(* IEC 61131-3 sources: daoli-st-library/DL_Process (part 38) *)

(* ---- FB_DL_InlineCheckweighGauge.st ---- *)
(*==============================================================================
 * 组件名称 (Component)  : FB_DL_InlineCheckweighGauge
 * 所属子库 (Sublibrary) : DL_Process
 * 当前版本 (Version)    : 1.0.0
 * 兼容性 (Platform)     : CODESYS 3.5 / TwinCAT 3 / 汇川 InoProShop（纯标准元素，无方言）
 * 功能描述 (Function)   : 在线称重动态窗判据与 σ 控制图。逐件判欠重/超重（不平顺：平滑会
 *                         漏掉单件超重），滑动统计窗给均值与样本标准差（分母 n−1，n≥5 前置
 *                         保证防除零），满窗后才判 σ 越控制限；可选的 ±3σ 冲击剔除只影响
 *                         统计窗，不影响逐件判据。不做传感器标定、不做零点跟踪（另有专件）、
 *                         不做剔除机构驱动。
 * 溯源 (Origin)         : 道莅 clean-room 防御性实现
 * 本文件内含 (Contains) : TYPE E_DL_GaugeWin / FUNCTION_BLOCK FB_DL_InlineCheckweighGauge
 * 依赖 (Depends)        : 无（仅 Standard.library 的 SQRT / ABS / MIN）
 * 红线自检 (Redline)    : 无外部全局变量、无硬件地址直引 ｜ 全变量中英双语同行注释
 *                         公差与控制限判零防除零 ｜ 样本非有限即丢弃并计丢弃数 ｜ 标准差前置
 *                         n≥5 且分母 n−1 ｜ σ 仅满窗判 ｜ 枚举显式赋值 ｜ CASE 含 ELSE 兜底
 *                         ｜ 本件无定时器/沿实例，全部为周期算术，故无周期刷新项
 * 错误码表 (Codes)      : 16#0005_0444 就绪（窗口统计正常）
 *                         16#0005_0445 预留：本版不发码（下一轮区间起点，禁止回填）
 *                         16#0005_0446 故障级 组态非法（公差 ≤0、窗长 <5、σ 限 ≤0）
 *                         16#0005_0447 故障级 目标重量非有限（逐件判据停判，统计继续）
 *                         16#0005_0448 信息级 样本非有限已丢弃（计入丢弃数）
 * 修订历史 (Revision)   : 2026-11-17  v1.0.0  首版入库 · R28 · 阶段三批 4
 * 验收向量 (Acceptance) : 正向 目标 500 g、公差 ±5、10 件 500±1 → 均值 ≈500、σ ≈0.7、
 *                         无报警
 *                         反向 一件 508 g → bOver 单件置位、uRejectCnt 不增（非剔除开关）、
 *                         均值仍 ≈500；σ 升到 6 超控制限 2 → bSpcAlarm；样本给 NaN →
 *                         16#0005_0448 且丢弃数 +1；窗长给 3 → 16#0005_0446
 *============================================================================*)

(*-----------------------------------------------------------------------------
 * 枚举: E_DL_GaugeWin（归属本功能块，同文件发布，全库唯一定义）
 *----------------------------------------------------------------------------*)
TYPE E_DL_GaugeWin :
(
    eEmpty := 0,    // 空窗：尚无有效样本 / Empty window, no valid sample yet
    eFill  := 10,   // 填充中：样本数未满窗长 / Filling, the sample count is below the window length
    eFull  := 20,   // 满窗：均值与 σ 可信 / Full window, the mean and sigma are trustworthy
    eFault := 99    // 故障：组态非法 / Fault, the configuration is invalid
);
END_TYPE

FUNCTION_BLOCK FB_DL_InlineCheckweighGauge
VAR_INPUT
    bEnable        : BOOL := FALSE;       // 使能 / Enable
    bSampleValid   : BOOL := FALSE;       // 本拍有有效样本 / A valid sample is present in this scan
    fWeight_g      : REAL := 0.0;         // 件重 [g]，域 0~50000 / Piece weight in grammes, domain 0 to 50000
    fTarget_g      : REAL := 500.0;       // 目标重量 [g] / Target weight in grammes
    fTolUp_g       : REAL := 5.0;         // 上公差带 [g]，须 >0 / Upper tolerance in grammes, must be positive
    fTolLow_g      : REAL := 5.0;         // 下公差带 [g]，须 >0 / Lower tolerance in grammes, must be positive
    uWinSamples    : UINT := 10;          // 统计窗长 [个]，域 5~50 / Statistical window length, domain 5 to 50
    fSigmaLimit_g  : REAL := 2.0;         // σ 控制限 [g]，域 0.1~20 / Sigma control limit in grammes, domain 0.1 to 20
    bOutlierReject : BOOL := FALSE;       // ±3σ 冲击剔除开关 / Plus minus three sigma outlier rejection switch
END_VAR
VAR_OUTPUT
    fMeanOut_g     : REAL;                // 窗口均值 [g] / Window mean in grammes
    fSigmaOut_g    : REAL;                // 窗口标准差 [g] / Window standard deviation in grammes
    bUnder         : BOOL;                // 本件欠重（逐件判据） / This piece is underweight
    bOver          : BOOL;                // 本件超重（逐件判据） / This piece is overweight
    bSpcAlarm      : BOOL;                // σ 越控制限（满窗后才判） / Sigma above the control limit, judged on a full window only
    uRejectCnt     : UDINT;               // 剔除件数 [件]（±3σ 剔除） / Outlier rejection count
    uSpcCnt        : UDINT;               // SPC 越限次数 [次] / SPC limit violation count
    eErr           : UDINT;               // 错误码，段位 16#0005_xxxx / Error code in segment 16#0005_xxxx
END_VAR
VAR
    _eWin          : E_DL_GaugeWin := E_DL_GaugeWin.eEmpty; // 窗口相位 / Window phase
    _bInit         : BOOL := FALSE;       // 首扫标志，取非判定 / First-scan flag, tested negated
    _bCfgOk        : BOOL;                // 组态合法标志 / Configuration valid flag
    _bTgtOk        : BOOL;                // 目标有限标志 / Target finite flag
    _bSpcLatched   : BOOL := FALSE;       // SPC 报警锁存（单拍计数用） / SPC alarm latch for one-shot counting
    _uWinEff       : UINT := 10;          // 生效窗长（钳制后）[个] / Effective window length after clamping
    _uIdx          : UINT := 1;           // 环形写指针 / Circular write index
    _uFill         : UINT := 0;           // 已填样本数 [个] / Number of samples collected
    _fSum          : REAL := 0.0;         // 样本和 [g] / Sample sum
    _fMean         : REAL := 0.0;         // 窗口均值 [g] / Window mean
    _fMeanOut_g    : REAL := 0.0;         // 窗口均值中间量（出口映射源）[g] / Window mean intermediate, source of the outlet [g]
    _fVar          : REAL := 0.0;         // 样本方差 [g²] / Sample variance
    _afWin         : ARRAY[1..50] OF REAL; // 样本环形窗 [g] / Sample ring buffer
    _iLoop         : INT;                 // 统计循环索引 / Statistical loop index
    _iGuard        : INT;                 // 防死循环计数器 / Loop guard counter
END_VAR
VAR CONSTANT
    DL_CW_READY    : UDINT := 16#0005_0444;  // 就绪码 / Ready code
    DL_CW_CFG_BAD  : UDINT := 16#0005_0446;  // 故障级组态非法码 / Fault code for bad configuration
    DL_CW_TGT_BAD  : UDINT := 16#0005_0447;  // 故障级目标非有限码 / Fault code for a non-finite target
    DL_CW_SKIP     : UDINT := 16#0005_0448;  // 信息级样本丢弃码 / Info code for a discarded sample
    DL_CW_WIN_LO   : UINT := 5;              // 窗长下限 [个] / Window length lower bound
    DL_CW_WIN_HI   : UINT := 50;             // 窗长上限 [个] / Window length upper bound
    DL_CW_SIG_LO   : REAL := 0.1;            // σ 控制限下限 [g] / Sigma limit lower bound
    DL_CW_SIG_HI   : REAL := 20.0;           // σ 控制限上限 [g] / Sigma limit upper bound
    DL_CW_LOOP_MAX : INT := 60;              // 循环保护上限 / Loop guard bound
    DL_CW_EPS      : REAL := 1.0E-6;         // 浮点判零容差 / Float zero tolerance
END_VAR

// 段 1｜输出与单拍标志预置
bUnder := FALSE;                                    // 欠重预清 / Underweight pre-cleared
bOver := FALSE;                                     // 超重预清 / Overweight pre-cleared
bSpcAlarm := FALSE;                                 // SPC 报警预清 / SPC alarm pre-cleared
eErr := 0;                                          // 错误码预清 / Error code pre-cleared

// 段 2｜首扫初始化（判据取非，R19）
IF NOT _bInit THEN
    _afWin[1] := 0.0;                               // 环形窗首元素预置 [g] / Ring buffer first element pre-set
    _eWin := E_DL_GaugeWin.eEmpty;                  // 窗口相位起点 / Window phase starts empty
    _bInit := TRUE;                                 // 首扫只做一次 / The first scan runs once
END_IF

// 段 3｜组态闸（公差与控制限判零防除零；窗长 <5 使 σ 不可信）
_bCfgOk := (fTolUp_g > 0.0) AND (fTolLow_g > 0.0)
        AND NOT ((fSigmaLimit_g <> fSigmaLimit_g) OR ((fSigmaLimit_g - fSigmaLimit_g) <> (fSigmaLimit_g - fSigmaLimit_g)))
        AND (fSigmaLimit_g >= DL_CW_SIG_LO) AND (fSigmaLimit_g <= DL_CW_SIG_HI)
        AND (uWinSamples >= DL_CW_WIN_LO) AND (uWinSamples <= DL_CW_WIN_HI);
_bTgtOk := NOT ((fTarget_g <> fTarget_g) OR ((fTarget_g - fTarget_g) <> (fTarget_g - fTarget_g)));
IF NOT _bCfgOk THEN
    eErr := DL_CW_CFG_BAD;                          // 故障级：组态非法 / Fault, bad configuration
    _eWin := E_DL_GaugeWin.eFault;
ELSE
    _uWinEff := uWinSamples;                        // 采用组态窗长 [个] / Use the configured window length
END_IF
IF NOT _bTgtOk THEN
    eErr := DL_CW_TGT_BAD;                          // 故障级：目标非有限（逐件判据停判） / Fault, the target is not finite
END_IF

// 段 4｜逐件判据（不平顺，单件即判；目标不可读时停判）
IF bEnable AND bSampleValid AND _bTgtOk THEN
    IF (fWeight_g <> fWeight_g) OR ((fWeight_g - fWeight_g) <> (fWeight_g - fWeight_g)) THEN
        eErr := DL_CW_SKIP;                         // 信息级：样本非有限，丢弃 / Info, the sample is not finite and is discarded
        uRejectCnt := uRejectCnt + 1;               // 丢弃计数 +1 [件] / Discard count incremented
    ELSE
        IF fWeight_g < (fTarget_g - fTolLow_g) THEN
            bUnder := TRUE;                         // 本件欠重 / This piece is underweight
        END_IF
        IF fWeight_g > (fTarget_g + fTolUp_g) THEN
            bOver := TRUE;                          // 本件超重 / This piece is overweight
        END_IF
        // 冲击剔除（±3σ，仅满窗且开关有效时；剔除只影响统计窗）
        IF bOutlierReject AND (_uFill >= DL_CW_WIN_LO) AND (fSigmaOut_g > DL_CW_EPS) THEN
            IF ABS(fWeight_g - _fMean) > (3.0 * fSigmaOut_g) THEN
                uRejectCnt := uRejectCnt + 1;       // ±3σ 剔除 +1 [件] / Outlier rejected
            ELSE
                _fSum := _fSum - _afWin[_uIdx];                 // 换出最旧样本 [g] / Remove the oldest sample
                _afWin[_uIdx] := fWeight_g;                     // 写入新样本 [g] / Insert the new sample
                _fSum := _fSum + fWeight_g;                     // 样本和更新 [g] / Update the sum
                _uIdx := _uIdx + 1;
                IF _uIdx > _uWinEff THEN
                    _uIdx := 1;                                 // 环形回卷 / Ring wrap
                END_IF
                IF _uFill < _uWinEff THEN
                    _uFill := _uFill + 1;                       // 已填样本数 +1 [个] / Sample count incremented
                END_IF
            END_IF
        ELSE
            _fSum := _fSum - _afWin[_uIdx];                     // 换出最旧样本 [g] / Remove the oldest sample
            _afWin[_uIdx] := fWeight_g;                         // 写入新样本 [g] / Insert the new sample
            _fSum := _fSum + fWeight_g;                         // 样本和更新 [g] / Update the sum
            _uIdx := _uIdx + 1;
            IF _uIdx > _uWinEff THEN
                _uIdx := 1;                                     // 环形回卷 / Ring wrap
            END_IF
            IF _uFill < _uWinEff THEN
                _uFill := _uFill + 1;                           // 已填样本数 +1 [个] / Sample count incremented
            END_IF
        END_IF
    END_IF
END_IF

// 段 5｜均值与样本标准差（分母 n−1，n≥5 前置保证防除零）
IF _uFill > 0 THEN
    _fMean := _fSum / UINT_TO_REAL(_uFill);         // 窗口均值 [g] / Window mean
END_IF
_fMeanOut_g := _fMean;                              // 均值出口 [g] / Mean output
_fVar := 0.0;                                       // 方差清零 [g²] / Variance reset
IF _uFill >= DL_CW_WIN_LO THEN
    _iLoop := 1;
    _iGuard := 0;
    WHILE (_iLoop <= UINT_TO_INT(_uWinEff)) AND (_iGuard < DL_CW_LOOP_MAX) DO
        _fVar := _fVar + ((_afWin[_iLoop] - _fMean) * (_afWin[_iLoop] - _fMean));   // 偏差平方累加 [g²] / Squared deviation accumulated
        _iLoop := _iLoop + 1;
        _iGuard := _iGuard + 1;                     // 防死循环计数 / Loop guard incremented
    END_WHILE
    _fVar := _fVar / UINT_TO_REAL(_uWinEff - 1);    // 样本方差（分母 n−1）[g²] / Sample variance with n minus one
    fSigmaOut_g := SQRT(_fVar);                     // 样本标准差 [g] / Sample standard deviation
ELSE
    fSigmaOut_g := 0.0;                             // 样本不足：σ 记 0（不参与判据） / Not enough samples, sigma reported as zero
END_IF

// 段 6｜σ 控制图（仅满窗判；越限只在锁存沿计数一次）
IF (_uFill >= _uWinEff) AND (_uWinEff >= DL_CW_WIN_LO) THEN
    IF fSigmaOut_g > fSigmaLimit_g THEN
        bSpcAlarm := TRUE;                          // σ 越控制限 / Sigma above the control limit
        IF NOT _bSpcLatched THEN
            uSpcCnt := uSpcCnt + 1;                 // 越限次数 +1（沿计数）[次] / Violation count incremented on the edge
            _bSpcLatched := TRUE;
        END_IF
    ELSE
        _bSpcLatched := FALSE;                      // 回限内：锁存解除 / Back inside the limit, the latch is released
    END_IF
END_IF

// 段 7｜窗口相位映射（ENUM + CASE + ELSE 兜底）
CASE _eWin OF
    E_DL_GaugeWin.eEmpty:
        IF _uFill > 0 THEN
            _eWin := E_DL_GaugeWin.eFill;           // 有样本：进入填充 / Samples exist, go filling
        END_IF
    E_DL_GaugeWin.eFill:
        IF _uFill >= _uWinEff THEN
            _eWin := E_DL_GaugeWin.eFull;           // 满窗 / Window full
        END_IF
    E_DL_GaugeWin.eFull:
        IF _uFill < _uWinEff THEN
            _eWin := E_DL_GaugeWin.eFill;           // 窗被重置 / The window was reset
        END_IF
    E_DL_GaugeWin.eFault:
        IF _bCfgOk THEN
            _eWin := E_DL_GaugeWin.eEmpty;          // 组态修正：回空窗 / Configuration fixed, back to empty
        END_IF
        eErr := DL_CW_CFG_BAD;                      // 故障级：组态非法保持 / Fault, the configuration error is held
    ELSE
        // 非法相位兜底（故障级）
        eErr := DL_CW_CFG_BAD;
        _eWin := E_DL_GaugeWin.eFault;
END_CASE
IF eErr = 0 THEN
    eErr := DL_CW_READY;                            // 无事件回就绪码 / Ready code when nothing else applies
END_IF
END_FUNCTION_BLOCK

(* ---- FB_DL_InvInsulTestSeq.st ---- *)
(*
  FB_DL_InvInsulTestSeq  —  逆变器绝缘测试加压-保持-泄放联锁顺控 / Inverter insulation test sequence with discharge interlock
  分类 Category : DL_Process
  码位 Code     : 16#06_0_98
  版本 Version  : 1.0.0
  溯源 Source   : ISA-88 相模型语义借鉴 · clean-room 实现，仅借分类/参数域/命名，未复制源码
  功能 Function : 1) 加压-保持-泄放三态顺控（复用 FB_DL_InterlockMatrix 联锁前置）；
                  2) 加压中急停立即转泄放相（安全侧打断）；
                  3) 泄放未确认前禁放行下工序；相完成仅在泄放反馈确认后置位。
  边界 Boundary : ① 泄放未确认前禁放行下工序（安全侧默认，bTestOk 不置位）；
                  ② 加压中急停立即转泄放相（打断优先级最高）；
                  ③ 各相超时独立 TON 升级；
                  ④ 测试电压反馈无效判「不可判」而非 OK；
                  ⑤ 输出三行同向：相状态 → 测试结论 → 联锁出口。
  依赖 Depends  : FB_DL_InterlockMatrix × 1（联锁前置，每拍无条件调用）

  码表 Error codes（本件子码步进 16#30 · 本格 98 与既有 9X 子码段冲突，错位至 C8/D8 避让）:
    16#0002_06C8 故障级：组态非法（任一相时长 <= 0 / 电压门限 <= 0）
    16#0002_06D8 故障级：相超时（加压/保持/泄放任一相在限时内未完成，锁存需复位）
    16#0002_06B8 信息级：电压反馈无效判不可判 / 泄放未确认不放行（不置 bError）
*)

TYPE E_DL_IitPhase :
(
    eIdle       := 0,  // 空闲 / Idle
    ePressurize := 10, // 加压相 / HV apply phase
    eHold       := 20, // 保持相 / Hold phase
    eDischarge  := 30, // 泄放相 / Discharge phase
    eDone       := 40, // 测试完成（泄放已确认）/ Test done, discharge confirmed
    eFault      := 90  // 超时/联锁故障锁定 / Timeout or interlock fault locked
);
END_TYPE

FUNCTION_BLOCK FB_DL_InvInsulTestSeq
VAR_INPUT
    bTestCmd      : BOOL;                           // 测试启动命令 / Test start command
    bEStop        : BOOL;                           // 急停（加压/保持相打断转泄放）/ Emergency stop
    bVoltFbOk     : BOOL;                           // 电压反馈有效前置 / Voltage feedback valid flag
    fVoltFb       : REAL;                           // 测试电压反馈 [V] / Test voltage feedback [V]
    fVoltSp       : REAL := 1000.0;                 // 测试电压设定 [V]，域 > 0 / Test voltage setpoint [V]
    fVoltWinV     : REAL := 50.0;                   // 保持相电压窗半宽 [V]，域 > 0 / Hold voltage window [V]
    bDischargeFb  : BOOL;                           // 泄放反馈（残压低于安全值）/ Discharge feedback, residual below safe
    bReset        : BOOL;                           // 复位，上升沿清故障 / Reset, clears fault
    tApplyMax     : TIME := T#10S;                  // 加压相限时 [s]，域 > 0 / Apply phase timeout
    tHoldMax      : TIME := T#5S;                   // 保持相限时 [s]，域 > 0 / Hold phase timeout
    tDischMax     : TIME := T#30S;                  // 泄放相限时 [s]，域 > 0 / Discharge phase timeout
    fEps          : REAL := 1.0E-6;                 // 浮点判零容差 [1] / Floating zero tolerance
END_VAR
VAR_OUTPUT
    bApplyHv      : BOOL;                           // 加压出口 / HV apply output
    bDischargeCmd : BOOL;                           // 泄放命令出口 / Discharge command output
    bTestOk       : BOOL;                           // 测试结论（仅在泄放确认后置位）/ Test verdict, only after discharge confirmed
    bInterlock    : BOOL;                           // 联锁出口（TRUE = 允许加压）/ Interlock output
    bIndeterminate: BOOL;                           // 不可判标志（反馈无效）/ Indeterminate flag
    bError        : BOOL;                           // 故障标志，与故障级码配对 / Fault flag
    uErrorId      : UDINT;                          // 事件码，0 = 无事件 / Event code
    eStateOut     : E_DL_IitPhase;                  // 状态机当前态，段尾单点映射 / Phase mapped at tail
END_VAR
VAR
    _eState       : E_DL_IitPhase := E_DL_IitPhase.eIdle;  // 内部状态 / Internal state
    fbIlk         : FB_DL_InterlockMatrix;          // 联锁矩阵实例（无条件调用）/ Interlock matrix instance
    rtrStart      : R_TRIG;                         // 启动沿 / Start edge
    rtrReset      : R_TRIG;                         // 复位沿 / Reset edge
    tonApply      : TON;                            // 加压相超时（独立 TON）/ Apply timeout
    tonHold       : TON;                            // 保持相超时 / Hold timeout
    tonDisch      : TON;                            // 泄放相超时 / Discharge timeout
    abCondOk      : ARRAY[0..15] OF BOOL;           // 联锁条件表 / Interlock condition table
    auInvertMask  : WORD;                           // 取反掩码 / Invert mask
    auTripMask    : WORD;                           // 停机级掩码 / Trip-class mask
    bCfgOk        : BOOL;                           // 组态合法标志 / Configuration valid
    bVoltOk       : BOOL;                           // 电压反馈本拍有效 / Voltage feedback valid
    bVoltInWin    : BOOL;                           // 保持相电压在窗 / Hold voltage in window
    bIlkPermit    : BOOL;                           // 联锁放行 / Interlock permit
    uFault        : UDINT;                          // 锁存故障码 / Latched fault code
    uInfo         : UDINT;                          // 信息级码 / Information code
END_VAR

(* === 段 0 · 实例刷新 === *)
rtrStart(CLK := bTestCmd);                        // 每拍刷新启动沿
rtrReset(CLK := bReset);                          // 每拍刷新复位沿

(* === 段 1 · 组态闸 === *)
bCfgOk := (TIME_TO_REAL(tApplyMax) > fEps) AND (TIME_TO_REAL(tHoldMax) > fEps)
          AND (TIME_TO_REAL(tDischMax) > fEps)    // 三相时长正域
          AND (fVoltSp > fEps) AND (fVoltWinV > fEps)   // 电压设定与窗正域
          AND (fVoltSp = fVoltSp) AND (fVoltWinV = fVoltWinV);  // NaN 自反
IF NOT bCfgOk THEN
    uFault := 16#0002_06C8;                       // 故障级：组态非法
END_IF
IF rtrReset.Q AND bCfgOk THEN
    uFault := 16#0000;                            // 复位沿清锁存（解除路径可达）
END_IF
uInfo := 16#0000;                                 // 信息码每拍清零

(* === 段 2 · 相超时定时器（独立 TON，相离开即断输入，R40）=== *)
tonApply(IN := (_eState = E_DL_IitPhase.ePressurize), PT := tApplyMax);   // 加压相超时
tonHold(IN := (_eState = E_DL_IitPhase.eHold), PT := tHoldMax);           // 保持相超时
tonDisch(IN := (_eState = E_DL_IitPhase.eDischarge), PT := tDischMax);    // 泄放相超时
IF tonApply.Q OR tonHold.Q OR tonDisch.Q THEN
    uFault := 16#0002_06D8;                       // 故障级：任一相超时（锁存，非死等）
END_IF

(* === 段 3 · 联锁矩阵（无条件调用：急停未触发 + 电压反馈有效 + 复位态）=== *)
abCondOk[0] := NOT bEStop;                        // 条件 0 = 急停未触发
abCondOk[1] := bVoltFbOk;                         // 条件 1 = 电压反馈有效
abCondOk[2] := bDischargeFb OR (_eState = E_DL_IitPhase.eIdle);   // 条件 2 = 初始无残压或空闲态
auInvertMask := 16#0000;                          // 不取反
auTripMask := 16#0007;                            // 三条件均停机级
fbIlk(abConditionOk := abCondOk,                  // 条件表
      auInvertMask := auInvertMask,               // 取反掩码
      auTripMask := auTripMask,                   // 停机级掩码
      bEnable := TRUE,                            // 矩阵恒使能（安全联锁语义由条件表与停机级掩码承载）
      bReset := rtrReset.Q);                      // 复位沿透传
bIlkPermit := fbIlk.bPermitToRun;                 // 联锁放行
bInterlock := bIlkPermit;                         // 联锁出口

(* === 段 4 · 电压反馈域闸与保持窗判定 === *)
bVoltOk := bVoltFbOk AND (fVoltFb = fVoltFb) AND (fVoltFb >= 0.0) AND (fVoltFb < 1.0E30);  // NaN 自反 + 非负域
bVoltInWin := bVoltOk AND (ABS(fVoltFb - fVoltSp) <= fVoltWinV + fEps);   // 保持相电压在窗
IF (_eState = E_DL_IitPhase.eHold) AND (NOT bVoltOk) THEN
    uInfo := 16#0002_06B8;                        // 信息级：电压反馈无效判不可判
END_IF
bIndeterminate := (NOT bVoltOk) AND ((_eState = E_DL_IitPhase.eHold)
                    OR (_eState = E_DL_IitPhase.ePressurize));   // 不可判标志（非 OK）

(* === 段 5 · 主状态机（ENUM + CASE，含 ELSE 兜底）=== *)
CASE _eState OF
E_DL_IitPhase.eIdle :
    bTestOk := FALSE;                             // 空闲未完成
    IF uFault <> 16#0000 THEN
        _eState := E_DL_IitPhase.eFault;          // 故障优先
    ELSIF rtrStart.Q AND bIlkPermit AND bCfgOk THEN
        _eState := E_DL_IitPhase.ePressurize;     // 联锁放行才进加压相
    END_IF

E_DL_IitPhase.ePressurize :
    bApplyHv := bIlkPermit AND (uFault = 16#0000);   // 加压出口（联锁+无故障门控）
    bDischargeCmd := FALSE;                       // 加压相不出泄放命令
    IF bEStop THEN
        _eState := E_DL_IitPhase.eDischarge;      // 急停立即转泄放相（打断优先级最高）
    ELSIF uFault <> 16#0000 THEN
        _eState := E_DL_IitPhase.eFault;          // 超时转故障
    ELSIF bVoltInWin THEN
        _eState := E_DL_IitPhase.eHold;           // 电压进窗转保持相
    END_IF

E_DL_IitPhase.eHold :
    bApplyHv := TRUE;                             // 保持相维持加压
    bDischargeCmd := FALSE;                       // 保持相不出泄放命令
    IF bEStop THEN
        _eState := E_DL_IitPhase.eDischarge;      // 急停立即转泄放相
    ELSIF uFault <> 16#0000 THEN
        _eState := E_DL_IitPhase.eFault;          // 超时转故障
    ELSIF tonHold.Q THEN
        _eState := E_DL_IitPhase.eDischarge;      // 保持时限到转泄放相（正常流程）
    END_IF

E_DL_IitPhase.eDischarge :
    bApplyHv := FALSE;                            // 泄放相撤加压
    bDischargeCmd := TRUE;                        // 泄放命令保持
    IF uFault <> 16#0000 THEN
        _eState := E_DL_IitPhase.eFault;          // 泄放超时转故障
    ELSIF bDischargeFb AND (NOT bEStop) THEN
        bTestOk := TRUE;                          // 泄放反馈确认：相完成仅此时置位
        _eState := E_DL_IitPhase.eDone;           // 转完成相
    ELSE
        uInfo := 16#0002_06B8;                    // 信息级：泄放未确认不放行
    END_IF

E_DL_IitPhase.eDone :
    bApplyHv := FALSE;                            // 完成相撤加压
    bDischargeCmd := FALSE;                       // 完成相撤泄放命令
    bTestOk := TRUE;                              // 结论保持（防同拍抹除）
    IF rtrStart.Q THEN
        bTestOk := FALSE;                         // 新启动沿重开
        _eState := E_DL_IitPhase.ePressurize;     // 回加压相
    END_IF

E_DL_IitPhase.eFault :
    bApplyHv := FALSE;                            // 故障相撤加压
    bDischargeCmd := TRUE;                        // 故障安全侧：泄放命令保持
    bTestOk := FALSE;                             // 故障不出结论
    IF uFault = 16#0000 THEN
        _eState := E_DL_IitPhase.eIdle;           // 解锁回空闲
    END_IF

ELSE
    _eState := E_DL_IitPhase.eFault;              // 非法状态拦截
    uFault := 16#0002_06C8;                       // 故障级：相 ID 越界复用组态码段
END_CASE

(* === 段 6 · 输出映射 === *)
bError := (uFault <> 16#0000);                    // 故障标志仅由故障级码置位（R45 配对）
IF bError THEN
    uErrorId := uFault;                           // 故障级优先上报
ELSE
    uErrorId := uInfo;                            // 否则上报信息级码
END_IF
eStateOut := _eState;                             // 输出枚举段尾单点映射（N2 规则）
END_FUNCTION_BLOCK

(* ---- FB_DL_IvCurveScan.st ---- *)
(*
  FB_DL_IvCurveScan  —  IV 曲线扫描与特征点提取（Voc / Isc / FF + 扫描窗） / IV curve scan with Voc, Isc and fill-factor extraction inside a scan window
  分类 Category : DL_Process
  版本 Version  : 1.0.1
  来源 Source   : roadmap-pv-p1 — 光伏组件 IV 扫描测试工站真缺口
  溯源 Origin   : 道莅 clean-room 实现；Voc/Isc/Pmax/FF 为公开光伏特性参数定义式，未复制任何源码行
  功能 Function : 1) 扫描窗 eScan 内逐周期摄取 (fVmeasV, fImeasA) 采样：Voc = 电压最大值、
                  Isc = 电流最大值、Pmax = max(V×I) 功率最大值、nSample 采样计数；
                  2) 段 0 每拍单次求解 FF = Pmax/(Voc×Isc)，内核为纯计算子函数
                  FC_DL_IvFillFactorCalc（分母 <= 1.0E-9 返回 -1.0 哨兵，不饱和、不置 0），
                  判据与出口共用同一当拍量 _fFfPu，全件不存在同一子函数同参二次调用；
                  3) FF 低于 fFfMinPu 判组件异常（归因 eFfLow）；
                  4) 故障级单码 03A2，归因由 eCause 独立成员承载（R190）；
                  5) 信息级 04CA = 扫描完成沿；6) 解除式全当拍量（R240）。
  接口 Interface: 输入逐样电压/电流/扫描窗/最小采样数/FF 下限/电压量程；输出 Voc/Isc/Pmax/FF/采样数/码
  边界 Boundary : ① 组态闸：tScan <= T#0S、nSampleMin = 0、fFfMinPu <= 0.0、fVmaxV <= 0.0
                  任一成立 → 03A2 锁存；fFfMinPu / fVmaxV 同时做 NaN 自反判，否则 NaN 参与
                  `<= 0.0` 判据恒假 → 组态闸与「FF 越下限」判据双双静默失效；
                  ② 非有限输入（NaN 自反 + Inf 差值自减双判）→ 03A2 锁存且该样点不参与极值更新；
                  ③ 除零防护在子函数内前置判（分母非法返回 -1.0 哨兵，不饱和、不置 0）；
                  ④ 采样极值仅扫峰不回落（扫描窗内单调保持），窗口结束由 TON 单点置位；
                  ⑤ 扫描 TON / R_TRIG 段 0 无条件周期调用，IN 由相位派生；
                  ⑥ 零全局耦合（无 GVL / 无 VAR_EXTERNAL / 无直接物理地址访问）；
                  ⑦ 复位沿作用域（R283 返修）：eFault 相内 = 清故障三件 + 净重装窗内量并回 eIdle；
                  非故障相 = 仅清故障锁存三件，窗内量与相位一律不动；窗内量唯一重置点 =
                  eIdle→eScan 迁移（段 5），保证「复位不清窗」与「tonScan 不重装」自洽；
                  ⑧ 〔例外〕NaN 自反判 [x <> x] 与 Inf 差值自减判 [(x-x) <> (x-x)] 是浮点判等
                  禁令的唯一合法例外（R79），只许用于「非有限检测」；机检 G6 已对自反式加白名单。
  依赖 Depends  : Standard.library（TON / R_TRIG）
  码表 Error codes（Process 段 0005，故障窗口 03A2 / 信息窗口 04CA）:
    16#0005_03A2 故障级：IV 扫描故障总码（组态非法 / 输入非有限 / 采样数不足 / FF 越下限），
                 锁存至 bReset 上升沿；归因见 eCause，不新增码位（派单硬约束单码）
    16#0005_04CA 信息级：扫描完成沿（进入 eDone 单拍）
  修订历史 Revision :
    2026-11-19  v1.0.0  R43 首版（批次 2 · 序号 6）
    2026-11-19  v1.0.1  R45 返修（R283）：复位沿按相分域，非故障相不再清窗内极值与采样计数
                        （曾致 eScan 中复位后半窗从零累积、与 tonScan 不重装自相矛盾）；
                        FF 计算上移段 0 单次求解 _fFfPu，段 3 判据与 eEval 相改读当拍量，
                        删除同一 FC 同参双调用；出口 fFfPu 恒等 _fFfPu，消除 eDone 相 FF 恒 0；
                        组态闸补 NaN 自反判；边界新增⑦⑧；引脚契约零变更（PATCH）
*)

TYPE E_DL_IvsState :
(
    eIdle  := 0,      // 未使能待启动 / Idle, waiting start
    eScan  := 10,     // 扫描窗内逐样摄取 / Sampling inside scan window
    eEval  := 20,     // 特征点求解与判据 / Feature evaluation
    eDone  := 50,     // 扫描完成 / Done
    eFault := 90      // 故障锁存相 / Fault latched phase
);
END_TYPE

TYPE E_DL_IvsCause :
(
    eNone       := 0, // 无故障成因 / No cause
    eCfgIllegal := 1, // 组态非法 / Illegal configuration
    eNonFinite  := 2, // 输入非有限 / Non-finite input
    eSampleFew  := 3, // 采样数不足 / Too few samples
    eFfLow      := 4  // FF 越下限（含分母不可计算时 FF 不可达下限） / Fill factor below limit
);
END_TYPE

FUNCTION FC_DL_IvFillFactorCalc : REAL
VAR_INPUT
    fPmaxW : REAL;    // 最大功率 [W] / Maximum power
    fVocV  : REAL;    // 开路电压 [V] / Open-circuit voltage
    fIscA  : REAL;    // 短路电流 [A] / Short-circuit current
END_VAR
(* 纯计算子函数：FF = Pmax / (Voc × Isc)；分母 <= 1.0E-9 返回 -1.0 哨兵（不饱和、不置 0） *)
IF (fVocV <= 1.0E-9) OR (fIscA <= 1.0E-9) THEN      // 除零前置判（分母正域检查） / Divide-by-zero guard
    FC_DL_IvFillFactorCalc := -1.0;                 // 哨兵：分母非法 / Sentinel for invalid denominator
ELSE
    FC_DL_IvFillFactorCalc := fPmaxW / (fVocV * fIscA);   // 填充因子（无量纲） / Fill factor
END_IF
END_FUNCTION

FUNCTION_BLOCK FB_DL_IvCurveScan
VAR_INPUT
    fVmeasV      : REAL := 0.0;       // 逐样电压 [V] / Per-sample voltage
    fImeasA      : REAL := 0.0;       // 逐样电流 [A] / Per-sample current
    tScan        : TIME := T#2S;      // 扫描窗时长 [ms]，域 > 0 / Scan window duration
    nSampleMin   : UDINT := 20;       // 最小采样点数 [点]，域 > 0 / Minimum sample count
    fFfMinPu     : REAL := 0.60;      // FF 下限 [p.u.]，域 > 0 / Fill factor lower limit
    fVmaxV       : REAL := 60.0;      // 电压量程上限 [V]，域 > 0 / Voltage range limit
    bStart       : BOOL := FALSE;     // 启动命令（电平）[-] / Start command
    bReset       : BOOL := FALSE;     // 复位命令，上升沿清故障 [-] / Reset edge
END_VAR
VAR_OUTPUT
    eState       : E_DL_IvsState;     // 状态出口，段 6 单点映射 / State outlet
    eCause       : E_DL_IvsCause;     // 故障成因出口（R190） / Fault cause outlet
    fVocV        : REAL;              // 开路电压 [V] / Open-circuit voltage
    fIscA        : REAL;              // 短路电流 [A] / Short-circuit current
    fPmaxW       : REAL;              // 最大功率 [W] / Maximum power
    fFfPu        : REAL;              // 填充因子 [p.u.] / Fill factor
    nSampleCount : UDINT;             // 本次扫描采样点数 [点] / Sample count
    bCycleDone   : BOOL;              // 扫描完成标志 [-] / Scan done flag
    bError       : BOOL;              // 故障锁存标志 [-] / Fault latch flag
    nErrId       : UDINT;             // 事件码，0 = 无事件 / Event code
END_VAR
VAR
    _eState      : E_DL_IvsState := E_DL_IvsState.eIdle;   // 内部相位（CASE 唯一写入目标） / Internal phase
    _eCause      : E_DL_IvsCause := E_DL_IvsCause.eNone;   // 故障成因锁存（锁存量） / Latched cause
    tonScan      : TON;               // 扫描窗计时，每周期无条件调用 / Scan window timer
    rtReset      : R_TRIG;            // 复位沿实例，每周期无条件调用 / Reset edge
    _fVocV       : REAL;              // 扫描期电压极值（窗内保持） / Voltage peak held in window
    _fIscA       : REAL;              // 扫描期电流极值（窗内保持） / Current peak held in window
    _fPmaxW      : REAL;              // 扫描期功率极值（窗内保持） / Power peak held in window
    _nSample     : UDINT;             // 采样计数（窗内累计） / Sample counter
    _fPowW       : REAL;              // 当拍功率 [W] / Instantaneous power
    _fFfPu       : REAL;              // FF 当拍量 [p.u.]（段 0 单次求解，供判据与出口） / FF per-scan value
    _bNonFin     : BOOL;              // 输入非有限当拍量 [-] / Non-finite input flag
    _bCfgBad     : BOOL;              // 组态非法当拍量 [-] / Config illegal
    _bFault      : BOOL;              // 故障锁存位（锁存量） / Latched fault bit
    _uFault      : UDINT;             // 故障码锁存（锁存量） / Latched fault code
    _uInfo       : UDINT;             // 信息码，每拍重算 / Transient info code
END_VAR

(* —— 段 0：沿实例与定时器无条件周期刷新 + 非有限判定 + FF 单次求解 —— *)
_bNonFin := (fVmeasV <> fVmeasV) OR (fImeasA <> fImeasA)
         OR ((fVmeasV - fVmeasV) <> (fVmeasV - fVmeasV))
         OR ((fImeasA - fImeasA) <> (fImeasA - fImeasA));       // NaN 自反 + Inf 差值自减双判（禁令唯一例外 R79） / NaN and Inf detection
_bCfgBad := (fFfMinPu <> fFfMinPu) OR (fVmaxV <> fVmaxV)         // 组态实数 NaN 自反判（禁令唯一例外 R79） / NaN self-test on config reals
         OR (tScan <= T#0S) OR (nSampleMin = 0) OR (fFfMinPu <= 0.0) OR (fVmaxV <= 0.0);   // 组态非法当拍量 / Config illegal
rtReset(CLK := bReset);                                         // 复位沿，每拍必调 / Reset edge
tonScan(IN := (_eState = E_DL_IvsState.eScan), PT := tScan);    // 扫描窗计时（IN 由相位派生，跨相自动复位 R228A/B） / Scan window timer
_fFfPu := FC_DL_IvFillFactorCalc(fPmaxW := _fPmaxW, fVocV := _fVocV, fIscA := _fIscA);   // FF 当拍量：段 0 单次求解，判据与出口共用 / FF solved once per scan

(* —— 段 1：单拍量预清零（锁存量与窗内极值保持量不入清单） —— *)
_uInfo := 16#0000_0000;            // 信息码每拍重算 / Info recomputed
fVocV := 0.0;                      // Voc 出口缺省 0 / Voc default
fIscA := 0.0;                      // Isc 出口缺省 0 / Isc default
fPmaxW := 0.0;                     // Pmax 出口缺省 0 / Pmax default
fFfPu := 0.0;                      // FF 出口缺省 0 / FF default
bCycleDone := FALSE;               // 完成标志缺省 FALSE / Done default
nErrId := 16#0000_0000;            // 事件码缺省无事件 / Event code default

(* —— 段 2：复位沿（按相分域，R283） + 组态域闸 —— *)
IF rtReset.Q THEN                                  // 复位沿（当拍量） / Reset edge
    _bFault := FALSE;                              // 清故障锁存位（锁存量） / Clear fault latch
    _uFault := 16#0000_0000;                       // 清故障锁存码（锁存量） / Clear fault code
    _eCause := E_DL_IvsCause.eNone;                // 清成因（锁存量） / Clear cause
    IF _eState = E_DL_IvsState.eFault THEN         // 仅故障相做净重装 / Clean re-arm only from fault
        _fVocV := 0.0;                             // 清窗内电压极值 / Clear voltage peak
        _fIscA := 0.0;                             // 清窗内电流极值 / Clear current peak
        _fPmaxW := 0.0;                            // 清窗内功率极值 / Clear power peak
        _nSample := 0;                             // 清采样计数 / Clear sample counter
        _eState := E_DL_IvsState.eIdle;            // 故障相迁出唯一路径 / Sole exit from fault
    END_IF
END_IF
IF _bCfgBad THEN                                   // 组态域闸 / Config gate
    _uFault := 16#0005_03A2;                       // 故障级：IV 扫描故障总码 / Process fault code
    _bFault := TRUE;                               // 锁存置位 / Latch set
    bError := TRUE;                                // 故障标志同拍置位（R45 配对） / Error flag set same scan
    _eCause := E_DL_IvsCause.eCfgIllegal;          // 归因：组态非法 / Cause: illegal config
END_IF
IF (NOT _bFault) AND _bNonFin THEN                 // 输入非有限（当拍量） / Non-finite input
    _uFault := 16#0005_03A2;                       // 故障级：IV 扫描故障总码 / Process fault code
    _bFault := TRUE;                               // 锁存置位 / Latch set
    bError := TRUE;                                // 故障标志同拍置位（R45 配对） / Error flag set same scan
    _eCause := E_DL_IvsCause.eNonFinite;           // 归因：非有限 / Cause: non-finite
END_IF

(* —— 段 3：采样数不足与 FF 越下限（判据当拍量 _fFfPu；仅在 eEval 相判） —— *)
IF (NOT _bFault) AND (_eState = E_DL_IvsState.eEval) AND (_nSample < nSampleMin) THEN
    _uFault := 16#0005_03A2;                       // 故障级：IV 扫描故障总码 / Process fault code
    _bFault := TRUE;                               // 锁存置位 / Latch set
    bError := TRUE;                                // 故障标志同拍置位（R45 配对） / Error flag set same scan
    _eCause := E_DL_IvsCause.eSampleFew;           // 归因：采样不足 / Cause: too few samples
END_IF
IF (NOT _bFault) AND (_eState = E_DL_IvsState.eEval) AND (_fFfPu < fFfMinPu) THEN
    (* 含哨兵 -1.0：分母不可计算（Voc 或 Isc 过小）时 FF 不可达下限，按安全侧判组件异常，
       故此处不设 `>= 0.0` 前置闸——该前置闸会造成 eEval 无迁出（R228B 同类缺陷） / Sentinel included: unreachable FF fails safe *)
    _uFault := 16#0005_03A2;                       // 故障级：IV 扫描故障总码 / Process fault code
    _bFault := TRUE;                               // 锁存置位 / Latch set
    bError := TRUE;                                // 故障标志同拍置位（R45 配对） / Error flag set same scan
    _eCause := E_DL_IvsCause.eEfLow;               // 归因：FF 越下限 / Cause: fill factor low
END_IF

(* —— 段 4：故障解除式（R240；全当拍量）：rtReset.Q / NOT _bCfgBad / NOT _bNonFin / NOT tonScan.Q ——
   解除式自证可满足（终审两式 1）：故障相内 _eState = eFault → tonScan.IN 恒假 → tonScan.Q 恒假；
   _bCfgBad 与 _bNonFin 由操作员/接线侧消除（组态改正、非有限输入消失），故四因子可同时为真，
   达式可满足、非 R152 恒假组合。 *)
IF rtReset.Q AND (NOT _bCfgBad) AND (NOT _bNonFin) AND (NOT tonScan.Q) THEN
    _bFault := FALSE;                              // 清故障锁存位（锁存量） / Clear fault latch
    _uFault := 16#0000_0000;                       // 清故障锁存码（锁存量） / Clear fault code
    _eCause := E_DL_IvsCause.eNone;                // 清成因（锁存量） / Clear cause
END_IF

(* —— 段 4A：故障锁存相位迁移闸 —— *)
IF _bFault AND (_eState <> E_DL_IvsState.eFault) THEN
    _eState := E_DL_IvsState.eFault;               // 锁存即入故障相 / Latch enters fault phase
END_IF

(* —— 段 5：相位机（CASE 全覆盖 + ELSE 兜底） —— *)
CASE _eState OF

E_DL_IvsState.eIdle:
    IF bStart AND (NOT _bFault) THEN           // 启动条件 / Start gate
        _fVocV := 0.0;                         // 窗内量唯一重置点（起扫） / Sole reset point of window peaks
        _fIscA := 0.0;                         // 清电流极值 / Reset current peak
        _fPmaxW := 0.0;                        // 清功率极值 / Reset power peak
        _nSample := 0;                         // 清采样计数 / Reset sample counter
        _eState := E_DL_IvsState.eScan;        // 进扫描相 / Enter scan
    END_IF

E_DL_IvsState.eScan:
    IF NOT _bNonFin THEN                                   // 仅有效样点参与极值（安全侧） / Valid samples only
        _nSample := _nSample + 1;                          // 采样计数递增 / Sample counter
        IF (fVmeasV > _fVocV) AND (fVmeasV <= fVmaxV) THEN
            _fVocV := fVmeasV;                             // 电压极值更新（量程钳制） / Voltage peak
        END_IF
        IF fImeasA > _fIscA THEN
            _fIscA := fImeasA;                             // 电流极值更新 / Current peak
        END_IF
        _fPowW := fVmeasV * fImeasA;                       // 当拍功率 / Instantaneous power
        IF _fPowW > _fPmaxW THEN
            _fPmaxW := _fPowW;                             // 功率极值更新 / Power peak
        END_IF
    END_IF
    IF tonScan.Q THEN                                      // 扫描窗到时（事件量） / Scan window elapsed
        _eState := E_DL_IvsState.eEval;                    // 进判据相 / Enter evaluation
    ELSIF NOT bStart THEN                                  // 撤启动（前置消失，R98 双出口） / Start released
        _eState := E_DL_IvsState.eIdle;                    // 回空闲（回 eIdle 时经 eIdle→eScan 才净重装） / Back to idle
    END_IF

E_DL_IvsState.eEval:
    IF _bFault THEN                                        // 段 3 已锁故障（含哨兵归因 eFfLow） / Fault already latched
        _eState := E_DL_IvsState.eFault;                   // 入故障相 / Enter fault phase
    ELSE                                                   // 分母合法且 FF 达下限 / Valid FF verdict
        _uInfo := 16#0005_04CA;                            // 信息级：扫描完成沿 / Info: scan complete edge
        _eState := E_DL_IvsState.eDone;                    // 进完成相 / Enter done
    END_IF

E_DL_IvsState.eDone:
    IF NOT bStart THEN                                     // 撤启动回空闲 / Start released returns idle
        _eState := E_DL_IvsState.eIdle;
    END_IF

E_DL_IvsState.eFault:
    ;                                                      // 故障相：仅段 4 复位沿可迁出 / Only reset exits

ELSE
    _uFault := 16#0005_03A2;                   // 故障级：非法相位兜底（归并总码） / Illegal phase fallback
    _bFault := TRUE;                           // 锁存置位 / Latch set
    bError := TRUE;                            // 故障标志同拍置位（R45 配对） / Error flag set same scan
    _eCause := E_DL_IvsCause.eCfgIllegal;      // 归因：相位非法归并组态 / Cause: phase illegal
    _eState := E_DL_IvsState.eFault;           // 强制回故障相 / Force fault phase

END_CASE

(* —— 段 6：出口单点映射（名实同源；锁存码回放） —— *)
fVocV := _fVocV;                               // Voc 出口 / Voc outlet
fIscA := _fIscA;                               // Isc 出口 / Isc outlet
fPmaxW := _fPmaxW;                             // Pmax 出口 / Pmax outlet
fFfPu := _fFfPu;                               // FF 出口 = 当拍量（eDone 相保持有效值） / FF from per-scan value
nSampleCount := _nSample;                      // 采样计数出口 / Sample count outlet
bCycleDone := (_eState = E_DL_IvsState.eDone); // 完成标志 / Done flag
IF _bFault THEN
    nErrId := _uFault;                         // 故障锁存码回放 / Replay latched code
    fFfPu := 0.0;                              // 故障相 FF 出口强制 0（安全侧，不输出哨兵） / FF forced zero in fault
ELSE
    nErrId := _uInfo;                          // 信息码 / Transient info
END_IF
bError := _bFault;                             // 故障标志同源 / Flag from latch
eState := _eState;                             // 状态出口 / State outlet
eCause := _eCause;                             // 成因出口 / Cause outlet

END_FUNCTION_BLOCK

(* ---- FB_DL_JiggerBatchRecipeSeq.st ---- *)
(*
  Name: FB_DL_JiggerBatchRecipeSeq
  Category: DL_Process
  Version: 1.0.0
  Round: R91 / 2026-11-25
  开源溯源：clean-room 自研（族 间歇式溢流染色与丝光整理，ST 开源生态实测 0 命中，无外部代码引入）
  功能：1) 染缸批次运行状态机，九相推进（含故障相）：
           待机 → 进布 → 进液 → 升温 → 保温 → 降温 → 水洗 → 出布 → （回待机）。
           待机相等 xStart 上升沿（必须边沿，防上电即在启动位自动进布）；
           进布相给进布命令等进布到位反馈；进液相开进液阀等液位达 fFillLevelMinPct；
           升温相开加热命令并把温度设定值置 fHeatTargetC，等温度达「目标 − 带宽」；
           保温相保持温度设定并计时 tHoldS；降温相开冷却命令、设定值置 fCoolTargetC，
           等温度降到「目标 + 带宽」；水洗相开进水阀等水洗到位反馈；
           出布相给出布命令等出布到位反馈，完成后置 xDone 锁存并回待机（保持到 xStart 撤下）。
        2) 步序跳转保护（本件的核心加固点）：状态机除判「本相完成条件」外，
           还必须复检「前相前置条件仍成立」，任一消失即锁码 0432 并进故障相：
           进液至水洗五相内 xLoadDoneFb 必须仍为 TRUE（布在缸内，防布卷被冲出）；
           升温至水洗五相内液位必须仍 >= fFillLevelMinPct（防干烧加热器与泵空转）。
           这是「跳步」（例如中途出布信号抖动）的唯一拦截位置。
        3) 每相独立超时 + 整序总超时：八个工作相各配「相定时 + 裕量」超时点，
           tonTotal 兜底整序总时长，九个超时源并发监视，任一命中即锁码进故障相。
  边界条件：1) 非有限值闸：温度、液位、目标温度、液位门槛、温度带宽、周期先过
           NOT(x > -DL_BIG AND x < DL_BIG)，同时拦 NaN 与 Inf；命中即锁码 0431 进故障相，
           绝不把 NaN 拿去与温度/液位阈比较（NaN 比较恒假会让到达条件永不成立且永不报错，R19）。
        2) 周期入参闸（R21）：本件不做斜率运算，fCycleS 仅作观测记录；
           非法周期改用缺省 DL_CYCLE_DEF = 0.1 s，并在组态闸中一并锁码 0431（同码归因，成员分离）。
        3) 阈值域闸：-DL_T_SPAN < fCoolTargetC < fHeatTargetC <= DL_T_SPAN、fTempBandK > DL_EPS、
           0.0 < fFillLevelMinPct <= DL_PCT_HI，越域锁码 0431
           （降温目标高于升温目标会让温度判据永不成立）。
        4) 单点赋值（R26）：六个命令位、温度设定、xDone / xBusy 全部在段 8 统一出口写一次，
           相位内只改 _eState / _fSpC / 锁存位，不在分支内各写一遍命令。
        5) 定时器周期刷新（R7）：十七个 TON 与两个边沿实例全部在 CASE 之外无条件调用，
           IN 由状态导出，相迁移即 IN 归假自复位（R188）。
        6) 故障解除路径：故障相内 xReset 上升沿 AND NOT xFault AND 入参/组态合法 → 清锁存回待机，
           回待机后必须重新给 xStart 上升沿才能再启动（不自恢复）。
        7) 状态机兜底：CASE 全态覆盖 + ELSE 强制回故障相并置码 0433、清全部输出。
        8) 输出安全初值（R25）：六个命令位初值 FALSE（失电即安全侧：不进液、不加热、不出布）；
           温度设定初值 = 实测温度（无升降温需求）。
           故障侧语义（R191 显式声明）：故障相 fTempSpC 优先冻结在实测温度 fTempC（有限值时），
           实测非有限则回落到已过二阶终闸的安全设定值，绝不把 NaN 传给下游；不给加热指令也不给
           强冷指令；xBusy := FALSE（降级置标志而不静默）。
  量纲自证：fTempC / fHeatTargetC / fCoolTargetC 为 [degC]，fTempBandK 为温差不 [K]，degC 差值以 K 计；
           fLevelPct / fFillLevelMinPct 为液位百分数 [%]，比较两侧同量纲；
           所有时间引脚为 [TIME]，相超时点 = [TIME] + [TIME] = [TIME]，与 TON 的 PT 同量纲。
  码表 Error codes（本件子带 0091_042x / 043x，故障级一律 3 行内置 _uFault/_bFault/_eState）:
    16#0091_0421 信息级：进布相等待进布到位反馈（不置故障位）
    16#0091_0422 故障级：进布相超时
    16#0091_0423 故障级：进液相超时（液位未达门槛）
    16#0091_0424 故障级：升温相超时（未达目标温度带）
    16#0091_0425 故障级：保温相超时
    16#0091_0426 故障级：降温相超时（未达降温目标带）
    16#0091_0427 故障级：水洗相超时
    16#0091_0428 故障级：出布相超时
    16#0091_0429 故障级：整序总超时
    16#0091_0430 故障级：外部故障输入 xFault
    16#0091_0431 故障级：入参非有限，或温度/液位/周期组态越域
    16#0091_0432 故障级：步序跳转保护（布不在缸内或液位不足，前置条件中途消失）
    16#0091_0433 故障级：状态机落 ELSE 兜底（非法相位 ID）
    16#0091_0434 信息级：批次完成保持中，等待撤令（不置故障位）

  修订历史 Revision :
    2026-11-25  v1.0.0  R91 首版
*)

TYPE E_DL_JbsBatchState :
(
    eJbsBatchIdle   := 0,     // 待机：等启动上升沿，全命令撤销 / Idle, awaiting start, all commands dropped
    eJbsBatchLoad   := 10,    // 进布：给进布命令等到位 / Loading, awaiting the load-done feedback
    eJbsBatchFill   := 20,    // 进液：开进液阀等液位 / Filling, awaiting the level threshold
    eJbsBatchHeat   := 30,    // 升温：开加热等目标温度带 / Heating, awaiting the target band
    eJbsBatchHold   := 40,    // 保温：保持温度设定并计时 / Holding, setpoint kept and timer running
    eJbsBatchCool   := 50,    // 降温：开冷却等降温目标带 / Cooling, awaiting the cool-down band
    eJbsBatchRinse  := 60,    // 水洗：开进水阀等水洗到位 / Rinsing, awaiting the rinse-done feedback
    eJbsBatchUnload := 70,    // 出布：给出布命令等到位 / Unloading, awaiting the unload-done feedback
    eJbsBatchFault  := 90     // 故障：锁存待解除 / Fault, latched awaiting release
);
END_TYPE

FUNCTION_BLOCK FB_DL_JiggerBatchRecipeSeq
VAR_INPUT
    xStart          : BOOL;    // 批次启动指令（上升沿有效）[bool] / Batch start command, edge triggered [bool]
    xReset          : BOOL;    // 故障复位（上升沿有效）[bool] / Fault reset, rising edge [bool]
    xFault          : BOOL;    // 外部故障汇总 [bool] / External fault aggregate [bool]
    xLoadDoneFb     : BOOL;    // 进布到位反馈 [bool] / Load-done feedback [bool]
    xFillDoneFb     : BOOL;    // 进液完成反馈（液位开关）[bool] / Fill-done feedback, level switch [bool]
    xRinseDoneFb    : BOOL;    // 水洗到位反馈 [bool] / Rinse-done feedback [bool]
    xUnloadDoneFb   : BOOL;    // 出布到位反馈 [bool] / Unload-done feedback [bool]
    fTempC          : REAL;    // 染液实测温度 [degC] / Measured dye liquor temperature [degC]
    fLevelPct       : REAL;    // 染液液位百分数 [%] / Dye liquor level percentage [%]
    fFillLevelMinPct : REAL;   // 进液完成液位门槛 [%] / Fill level threshold [%]
    fHeatTargetC    : REAL;    // 升温目标温度 [degC] / Heating target temperature [degC]
    fCoolTargetC    : REAL;    // 降温目标温度 [degC] / Cooling target temperature [degC]
    fTempBandK      : REAL;    // 到温判定带宽 [K] / At-target band width [K]
    fCycleS         : REAL;    // 任务周期（观测用）[s] / Task cycle time, for observation [s]
    tLoadS          : TIME;    // 进布相设定时长 [TIME] / Loading phase duration [TIME]
    tFillS          : TIME;    // 进液相设定时长 [TIME] / Filling phase duration [TIME]
    tHeatS          : TIME;    // 升温相设定时长 [TIME] / Heating phase duration [TIME]
    tHoldS          : TIME;    // 保温相设定时长 [TIME] / Holding phase duration [TIME]
    tCoolS          : TIME;    // 降温相设定时长 [TIME] / Cooling phase duration [TIME]
    tRinseS         : TIME;    // 水洗相设定时长 [TIME] / Rinsing phase duration [TIME]
    tUnloadS        : TIME;    // 出布相设定时长 [TIME] / Unloading phase duration [TIME]
END_VAR
VAR_OUTPUT
    xLoadCmd        : BOOL;    // 进布命令（安全侧：故障时停）[bool] / Load command, fail-safe [bool]
    xFillValveCmd   : BOOL;    // 进液阀命令（安全侧：故障时关）[bool] / Fill valve command, fail-safe [bool]
    xHeatCmd        : BOOL;    // 加热命令（安全侧：故障时停）[bool] / Heating command, fail-safe [bool]
    xCoolCmd        : BOOL;    // 冷却命令（安全侧：故障时停）[bool] / Cooling command, fail-safe [bool]
    xRinseCmd       : BOOL;    // 水洗进水阀命令（安全侧：故障时关）[bool] / Rinse valve command, fail-safe [bool]
    xUnloadCmd      : BOOL;    // 出布命令（安全侧：故障时停）[bool] / Unload command, fail-safe [bool]
    fTempSpC        : REAL;    // 染液温度设定值 [degC] / Dye liquor temperature setpoint [degC]
    xDone           : BOOL;    // 批次完成保持位 [bool] / Batch complete held flag [bool]
    xBusy           : BOOL;    // 批次进行中 [bool] / Batch busy flag [bool]
    eState          : E_DL_JbsBatchState;   // 状态出口，段尾单点映射 / State outlet, single-point mapped
    nErrId          : UDINT;   // 事件码，0 = 无事件 / Event code, 0 = none
END_VAR
VAR
    tonLoad         : TON;     // 进布相正常定时 [TIME] / Loading phase timer
    tonLoadOv       : TON;     // 进布相超时定时 [TIME] / Loading phase overrun timer
    tonFill         : TON;     // 进液相正常定时 [TIME] / Filling phase timer
    tonFillOv       : TON;     // 进液相超时定时 [TIME] / Filling phase overrun timer
    tonHeat         : TON;     // 升温相正常定时 [TIME] / Heating phase timer
    tonHeatOv       : TON;     // 升温相超时定时 [TIME] / Heating phase overrun timer
    tonHold         : TON;     // 保温相正常定时 [TIME] / Holding phase timer
    tonHoldOv       : TON;     // 保温相超时定时 [TIME] / Holding phase overrun timer
    tonCool         : TON;     // 降温相正常定时 [TIME] / Cooling phase timer
    tonCoolOv       : TON;     // 降温相超时定时 [TIME] / Cooling phase overrun timer
    tonRinse        : TON;     // 水洗相正常定时 [TIME] / Rinsing phase timer
    tonRinseOv      : TON;     // 水洗相超时定时 [TIME] / Rinsing phase overrun timer
    tonUnload       : TON;     // 出布相正常定时 [TIME] / Unloading phase timer
    tonUnloadOv     : TON;     // 出布相超时定时 [TIME] / Unloading phase overrun timer
    tonTotal        : TON;     // 整序总超时定时 [TIME] / Whole-sequence total timeout timer
    rtStart         : R_TRIG;  // 启动上升沿检测 [bool] / Start rising edge detector
    rtReset         : R_TRIG;  // 复位上升沿检测 [bool] / Reset rising edge detector
    _eState         : E_DL_JbsBatchState := E_DL_JbsBatchState.eJbsBatchIdle;   // 内部相位（CASE 唯一写入目标）
    _eStatePrev     : E_DL_JbsBatchState := E_DL_JbsBatchState.eJbsBatchIdle;   // 上一拍相位快照（周期末更新）
    _fSpC           : REAL := 0.0;    // 内部温度设定值状态量 [degC] / Internal temperature setpoint [degC]
    _fCycleUseS     : REAL := 0.1;    // 实际使用的周期值 [s] / Cycle time actually used [s]
    _fHeatLowC      : REAL := 0.0;    // 升温到温下限（目标 − 带宽）[degC] / Heating arrival low bound [degC]
    _fCoolHighC     : REAL := 0.0;    // 降温到温上限（目标 + 带宽）[degC] / Cooling arrival high bound [degC]
    _bFinOk         : BOOL := FALSE;  // 实值入参有限性总闸结果 / Finiteness gate aggregate result
    _bCfgOk         : BOOL := FALSE;  // 温度/液位/周期组态域闸结果 / Configuration domain gate result
    _bActive        : BOOL := FALSE;  // 序激活（进布至出布七相之一）[bool] / Sequence active flag
    _bFabInDrum     : BOOL := FALSE;  // 布在缸内（步序保护用）[bool] / Fabric inside the drum, step guard
    _bLevelOk       : BOOL := FALSE;  // 液位达门槛（步序保护用）[bool] / Level above threshold, step guard
    _bStepGuardBad  : BOOL := FALSE;  // 步序跳转保护触发标志 [bool] / Step-guard violation flag
    _bDoneL         : BOOL := FALSE;  // 完成位锁存（跨相保持）[bool] / Done latch held across phases
    _bFault         : BOOL := FALSE;  // 故障锁存位 [bool] / Latched fault flag
    _iPhaseChg      : INT := 0;       // 本拍相位切换计数（观测用）[-] / Phase-change count this cycle [-]
    _uInfo          : UDINT := 16#0000_0000;   // 信息码，每拍重算 / Info code, recomputed every cycle
    _uFault         : UDINT := 16#0000_0000;   // 故障码锁存 / Latched fault code
END_VAR
VAR CONSTANT
    DL_EPS          : REAL := 1.0E-9;     // 数值零闸阈值 [-] / Numeric zero gate threshold [-]
    DL_BIG          : REAL := 1.0E12;     // 非有限值闸量级上限 [-] / Finiteness gate magnitude [-]
    DL_CYCLE_DEF    : REAL := 0.1;        // 缺省任务周期 [s] / Default task cycle time [s]
    DL_CYCLE_MIN    : REAL := 0.001;      // 周期合理下限 [s] / Cycle time reasonable low bound [s]
    DL_CYCLE_MAX    : REAL := 10.0;       // 周期合理上限 [s] / Cycle time reasonable high bound [s]
    DL_T_SPAN       : REAL := 300.0;      // 温度量级闸跨度 [degC] / Temperature magnitude gate span [degC]
    DL_PCT_HI       : REAL := 100.0;      // 液位百分数物理上限 [%] / Level percentage upper bound [%]
    DL_OVER_MARGIN  : TIME := T#30M;      // 相超时相对正常定时的裕量 [TIME] / Phase overrun margin [TIME]
    DL_TOTAL_MAX    : TIME := T#24H;      // 整序总超时上限 [TIME] / Whole-sequence total timeout [TIME]
END_VAR

(* —— 段 0：单拍量预清零（锁存量 _uFault/_bFault/_bDoneL/_fSpC/_eStatePrev 不入清单，R187①） —— *)
_uInfo := 16#0000_0000;                     // 信息码每拍重算 / Info code recomputed
_iPhaseChg := 0;                            // 相位切换计数每拍重算 / Phase-change counter recomputed
nErrId := 16#0000_0000;                     // 事件码缺省无事件 / Event code defaults to none
_bStepGuardBad := FALSE;                    // 步序保护标志每拍重算 / Step-guard flag recomputed

(* —— 段 1：非有限值闸与组态域闸（R19：不拿 NaN 去比较温度与液位） —— *)
_bFinOk := (fTempC > -DL_BIG) AND (fTempC < DL_BIG)
           AND (fLevelPct > -DL_BIG) AND (fLevelPct < DL_BIG)
           AND (fFillLevelMinPct > -DL_BIG) AND (fFillLevelMinPct < DL_BIG)
           AND (fHeatTargetC > -DL_BIG) AND (fHeatTargetC < DL_BIG)
           AND (fCoolTargetC > -DL_BIG) AND (fCoolTargetC < DL_BIG)
           AND (fTempBandK > -DL_BIG) AND (fTempBandK < DL_BIG)
           AND (fCycleS > -DL_BIG) AND (fCycleS < DL_BIG);
_bCfgOk := (fTempBandK > DL_EPS)                        // 温度带宽必须为正
           AND (fFillLevelMinPct > 0.0)                 // 液位门槛必须为正
           AND (fFillLevelMinPct <= DL_PCT_HI)          // 液位门槛不得超 100 %
           AND (fLevelPct >= 0.0) AND (fLevelPct <= DL_PCT_HI)      // 实测液位量级闸
           AND (fHeatTargetC > fCoolTargetC)            // 降温目标必须低于升温目标（方向固定）
           AND (ABS(fHeatTargetC) <= DL_T_SPAN)         // 目标温度量级闸
           AND (ABS(fCoolTargetC) <= DL_T_SPAN)         // 目标温度量级闸
           AND (ABS(fTempC) <= DL_T_SPAN)               // 实测温度量级闸
           AND (fCycleS >= DL_CYCLE_MIN) AND (fCycleS <= DL_CYCLE_MAX);

IF _bCfgOk THEN
    _fCycleUseS := fCycleS;                 // 合法周期原值使用（本件仅观测用）
ELSE
    _fCycleUseS := DL_CYCLE_DEF;            // 非法周期一律用缺省 0.1 s
END_IF

(* —— 段 2：派生态（激活、到温带、步序保护前置量） —— *)
_bActive := (_eState = E_DL_JbsBatchState.eJbsBatchLoad)
            OR (_eState = E_DL_JbsBatchState.eJbsBatchFill)
            OR (_eState = E_DL_JbsBatchState.eJbsBatchHeat)
            OR (_eState = E_DL_JbsBatchState.eJbsBatchHold)
            OR (_eState = E_DL_JbsBatchState.eJbsBatchCool)
            OR (_eState = E_DL_JbsBatchState.eJbsBatchRinse)
            OR (_eState = E_DL_JbsBatchState.eJbsBatchUnload);
_fHeatLowC := fHeatTargetC - fTempBandK;                                  // 升温到温下限 [degC]
_fCoolHighC := fCoolTargetC + fTempBandK;                                 // 降温到温上限 [degC]
_bFabInDrum := xLoadDoneFb;                                               // 布在缸内判据（反馈即状态）
_bLevelOk := _bFinOk AND _bCfgOk AND (fLevelPct >= fFillLevelMinPct);      // 液位达门槛判据

(* —— 段 3：步序跳转保护（R：前置条件中途消失即锁码，唯一拦截位置） —— *)
IF (NOT _bFault) THEN
    IF ((_eState = E_DL_JbsBatchState.eJbsBatchFill)
        OR (_eState = E_DL_JbsBatchState.eJbsBatchHeat)
        OR (_eState = E_DL_JbsBatchState.eJbsBatchHold)
        OR (_eState = E_DL_JbsBatchState.eJbsBatchCool)
        OR (_eState = E_DL_JbsBatchState.eJbsBatchRinse)) AND (NOT _bFabInDrum) THEN
        _bStepGuardBad := TRUE;             // 布已不在缸内：进液之后的相一律非法
    END_IF
    IF ((_eState = E_DL_JbsBatchState.eJbsBatchHeat)
        OR (_eState = E_DL_JbsBatchState.eJbsBatchHold)
        OR (_eState = E_DL_JbsBatchState.eJbsBatchCool)
        OR (_eState = E_DL_JbsBatchState.eJbsBatchRinse)) AND (NOT _bLevelOk) THEN
        _bStepGuardBad := TRUE;             // 液位不足：加热与循环相一律非法（防干烧）
    END_IF
END_IF

(* —— 段 4：定时器与边沿无条件周期刷新（R7：调用语句不得置于 IF/CASE 内） —— *)
rtStart(CLK := xStart);                                                                  // 启动上升沿，每拍必调
rtReset(CLK := xReset);                                                                  // 复位上升沿，每拍必调
tonLoad(IN := (_eState = E_DL_JbsBatchState.eJbsBatchLoad), PT := tLoadS);               // 进布相正常定时
tonLoadOv(IN := (_eState = E_DL_JbsBatchState.eJbsBatchLoad), PT := tLoadS + DL_OVER_MARGIN);        // 进布超时点
tonFill(IN := (_eState = E_DL_JbsBatchState.eJbsBatchFill), PT := tFillS);                // 进液相正常定时
tonFillOv(IN := (_eState = E_DL_JbsBatchState.eJbsBatchFill), PT := tFillS + DL_OVER_MARGIN);        // 进液超时点
tonHeat(IN := (_eState = E_DL_JbsBatchState.eJbsBatchHeat), PT := tHeatS);                // 升温相正常定时
tonHeatOv(IN := (_eState = E_DL_JbsBatchState.eJbsBatchHeat), PT := tHeatS + DL_OVER_MARGIN);        // 升温超时点
tonHold(IN := (_eState = E_DL_JbsBatchState.eJbsBatchHold), PT := tHoldS);                // 保温相正常定时
tonHoldOv(IN := (_eState = E_DL_JbsBatchState.eJbsBatchHold), PT := tHoldS + DL_OVER_MARGIN);        // 保温超时点
tonCool(IN := (_eState = E_DL_JbsBatchState.eJbsBatchCool), PT := tCoolS);                // 降温相正常定时
tonCoolOv(IN := (_eState = E_DL_JbsBatchState.eJbsBatchCool), PT := tCoolS + DL_OVER_MARGIN);        // 降温超时点
tonRinse(IN := (_eState = E_DL_JbsBatchState.eJbsBatchRinse), PT := tRinseS);             // 水洗相正常定时
tonRinseOv(IN := (_eState = E_DL_JbsBatchState.eJbsBatchRinse), PT := tRinseS + DL_OVER_MARGIN);     // 水洗超时点
tonUnload(IN := (_eState = E_DL_JbsBatchState.eJbsBatchUnload), PT := tUnloadS);          // 出布相正常定时
tonUnloadOv(IN := (_eState = E_DL_JbsBatchState.eJbsBatchUnload), PT := tUnloadS + DL_OVER_MARGIN);  // 出布超时点
tonTotal(IN := _bActive, PT := DL_TOTAL_MAX);                                             // 整序总超时

(* —— 段 5：全局故障拦截（优先级最高；已锁存则不再改写码值，禁同拍抹除） —— *)
IF xFault AND (NOT _bFault) THEN
    _uFault := 16#0091_0430;                // 故障级：外部故障输入
    _bFault := TRUE;                        // 锁存（3 行内置，R45 配对）
    _eState := E_DL_JbsBatchState.eJbsBatchFault;
END_IF
IF ((NOT _bFinOk) OR (NOT _bCfgOk)) AND (NOT _bFault) THEN
    _uFault := 16#0091_0431;                // 故障级：入参非有限或组态越域（内部成员已分离）
    _bFault := TRUE;                        // 锁存
    _eState := E_DL_JbsBatchState.eJbsBatchFault;
END_IF
IF _bStepGuardBad AND (NOT _bFault) THEN
    _uFault := 16#0091_0432;                // 故障级：步序跳转保护（前置条件中途消失）
    _bFault := TRUE;                        // 锁存
    _eState := E_DL_JbsBatchState.eJbsBatchFault;
END_IF
IF tonTotal.Q AND _bActive AND (NOT _bFault) THEN
    _uFault := 16#0091_0429;                // 故障级：整序总超时
    _bFault := TRUE;                        // 锁存
    _eState := E_DL_JbsBatchState.eJbsBatchFault;
END_IF

(* —— 段 6：相位机（只做迁移与设定值更新；出口在段 8 单点映射） —— *)
CASE _eState OF

E_DL_JbsBatchState.eJbsBatchIdle:
    _fSpC := fTempC;                        // 待机设定值跟随实测（无升降温需求，安全侧）
    IF NOT xStart THEN
        _bDoneL := FALSE;                   // 撤令即清完成位，为下一批重新武装
    ELSIF rtStart.Q AND _bFinOk AND _bCfgOk THEN
        _bDoneL := FALSE;                   // 新批次开始：清完成位（迁移前一次性清）
        _eState := E_DL_JbsBatchState.eJbsBatchLoad;          // 进进布相
    END_IF

E_DL_JbsBatchState.eJbsBatchLoad:
    _fSpC := fTempC;                        // 进布相不控温
    IF tonLoadOv.Q THEN
        _uFault := 16#0091_0422;            // 故障级：进布相超时
        _bFault := TRUE;                    // 锁存
        _eState := E_DL_JbsBatchState.eJbsBatchFault;
    ELSIF tonLoad.Q AND xLoadDoneFb THEN
        _eState := E_DL_JbsBatchState.eJbsBatchFill;          // 本拍合法事件优先于超时迁移（R275）
    ELSE
        _uInfo := 16#0091_0421;             // 信息级：等进布到位反馈（不置故障位）
    END_IF

E_DL_JbsBatchState.eJbsBatchFill:
    _fSpC := fTempC;                        // 进液相不控温
    IF tonFillOv.Q THEN
        _uFault := 16#0091_0423;            // 故障级：进液相超时
        _bFault := TRUE;                    // 锁存
        _eState := E_DL_JbsBatchState.eJbsBatchFault;
    ELSIF tonFill.Q AND _bLevelOk AND xFillDoneFb THEN
        _eState := E_DL_JbsBatchState.eJbsBatchHeat;          // 液位到：进升温相
    END_IF

E_DL_JbsBatchState.eJbsBatchHeat:
    _fSpC := fHeatTargetC;                  // 升温相设定值置升温目标
    IF tonHeatOv.Q THEN
        _uFault := 16#0091_0424;            // 故障级：升温相超时
        _bFault := TRUE;                    // 锁存
        _eState := E_DL_JbsBatchState.eJbsBatchFault;
    ELSIF tonHeat.Q AND (fTempC >= _fHeatLowC) THEN
        _eState := E_DL_JbsBatchState.eJbsBatchHold;          // 到温带：进保温相
    END_IF

E_DL_JbsBatchState.eJbsBatchHold:
    _fSpC := fHeatTargetC;                  // 保温相设定值保持在升温目标
    IF tonHoldOv.Q THEN
        _uFault := 16#0091_0425;            // 故障级：保温相超时
        _bFault := TRUE;                    // 锁存
        _eState := E_DL_JbsBatchState.eJbsBatchFault;
    ELSIF tonHold.Q THEN
        _eState := E_DL_JbsBatchState.eJbsBatchCool;          // 保温到点：进降温相
    END_IF

E_DL_JbsBatchState.eJbsBatchCool:
    _fSpC := fCoolTargetC;                  // 降温相设定值置降温目标
    IF tonCoolOv.Q THEN
        _uFault := 16#0091_0426;            // 故障级：降温相超时
        _bFault := TRUE;                    // 锁存
        _eState := E_DL_JbsBatchState.eJbsBatchFault;
    ELSIF tonCool.Q AND (fTempC <= _fCoolHighC) THEN
        _eState := E_DL_JbsBatchState.eJbsBatchRinse;         // 降到目标带：进水洗相
    END_IF

E_DL_JbsBatchState.eJbsBatchRinse:
    _fSpC := fCoolTargetC;                  // 水洗相保持降温目标（防回温）
    IF tonRinseOv.Q THEN
        _uFault := 16#0091_0427;            // 故障级：水洗相超时
        _bFault := TRUE;                    // 锁存
        _eState := E_DL_JbsBatchState.eJbsBatchFault;
    ELSIF tonRinse.Q AND xRinseDoneFb THEN
        _eState := E_DL_JbsBatchState.eJbsBatchUnload;        // 水洗到位：进出布相
    END_IF

E_DL_JbsBatchState.eJbsBatchUnload:
    _fSpC := fTempC;                        // 出布相不控温
    IF tonUnloadOv.Q THEN
        _uFault := 16#0091_0428;            // 故障级：出布相超时
        _bFault := TRUE;                    // 锁存
        _eState := E_DL_JbsBatchState.eJbsBatchFault;
    ELSIF tonUnload.Q AND xUnloadDoneFb THEN
        _bDoneL := TRUE;                    // 完成位锁存（跨相保持，段 8 单点映射）
        _eState := E_DL_JbsBatchState.eJbsBatchIdle;          // 回待机，完成位保持到撤令
    END_IF

E_DL_JbsBatchState.eJbsBatchFault:
    _fSpC := fTempC;                        // 故障相设定值冻结在实测（不给加热也不给强冷，R191 已声明）
    IF rtReset.Q AND (NOT xFault) AND _bFinOk AND _bCfgOk THEN
        _bFault := FALSE;                   // 解除路径：复位沿 + 外部故障消失 + 入参/组态合法（可达，R188）
        _uFault := 16#0000_0000;            // 清锁存码
        _bDoneL := FALSE;                   // 完成位一并清，避免故障后误报完成
        _eState := E_DL_JbsBatchState.eJbsBatchIdle;          // 回待机，需新上升沿才可再启动
    END_IF

ELSE
    _uFault := 16#0091_0433;                // 故障级：非法相位 ID 兜底
    _bFault := TRUE;                        // 锁存
    _bDoneL := FALSE;                       // 完成位清
    _fSpC := fTempC;                        // 兜底侧设定值冻结在实测
    _eState := E_DL_JbsBatchState.eJbsBatchFault;             // 强制回故障相

END_CASE

(* —— 段 7：后置段（相位快照与设定值域兜底） —— *)
IF _eState <> _eStatePrev THEN
    _iPhaseChg := _iPhaseChg + 1;           // 相位已切换：记一拍切换事件（观测用）
END_IF
_eStatePrev := _eState;                     // 快照在周期末尾统一更新
IF NOT (_fSpC > -DL_BIG AND _fSpC < DL_BIG) THEN
    _fSpC := fTempC;                        // 内部状态自检：非有限即回落实测值
END_IF
_fSpC := LIMIT(-DL_T_SPAN, _fSpC, DL_T_SPAN);   // 越量级钳制，防设定值发散
(* —— 段 7.5：LIMIT 后二阶终闸（R19 二阶形态）——
   LIMIT 对 NaN 会原样透传（内部比较全假走 ELSE 支），一次钳制不足以闸断通路，
   且上面那次回退源 fTempC 本身也可能非有限，故在钳制之后再判一次。 *)
IF NOT (_fSpC >= -DL_T_SPAN AND _fSpC <= DL_T_SPAN) THEN
    _fSpC := 0.0;                           // 双源皆非有限：0 degC 安全位 / Both sources non-finite: 0 degC safe
END_IF

(* —— 段 8：出口单点映射（名实同源；命令位由状态导出，故障侧一律撤销） —— *)
xLoadCmd := (_eState = E_DL_JbsBatchState.eJbsBatchLoad) AND (NOT _bFault);               // 进布命令
xFillValveCmd := (_eState = E_DL_JbsBatchState.eJbsBatchFill) AND (NOT _bFault);          // 进液阀
xHeatCmd := ((_eState = E_DL_JbsBatchState.eJbsBatchHeat)
             OR (_eState = E_DL_JbsBatchState.eJbsBatchHold)) AND (NOT _bFault);          // 加热：升温+保温
xCoolCmd := ((_eState = E_DL_JbsBatchState.eJbsBatchCool)
             OR (_eState = E_DL_JbsBatchState.eJbsBatchRinse)) AND (NOT _bFault);         // 冷却：降温+水洗
xRinseCmd := (_eState = E_DL_JbsBatchState.eJbsBatchRinse) AND (NOT _bFault);             // 水洗进水阀
xUnloadCmd := (_eState = E_DL_JbsBatchState.eJbsBatchUnload) AND (NOT _bFault);           // 出布命令
IF _bFault THEN
    IF (fTempC >= -DL_T_SPAN) AND (fTempC <= DL_T_SPAN) THEN
        fTempSpC := fTempC;                 // 故障侧优先回落实测温度（有限时保持原语义：冻结在实测）
    ELSE
        fTempSpC := _fSpC;                  // 实测非有限时回落到已过二阶终闸的安全值，绝不输出 NaN
    END_IF;
ELSE
    fTempSpC := _fSpC;                      // 正常侧设定值出口
END_IF
xDone := _bDoneL AND (NOT _bFault);                                                       // 完成位出口
xBusy := _bActive AND (NOT _bFault);                                                      // 进行中出口（故障时降级置假）
eState := _eState;                                                                        // 状态出口单点映射
IF _bFault THEN
    nErrId := _uFault;                      // 故障锁存码回放（不在故障相按当下输入重推断）
ELSIF _bDoneL THEN
    nErrId := 16#0091_0434;                 // 信息级：批次完成保持中，等待撤令
ELSE
    nErrId := _uInfo;                       // 信息码
END_IF

END_FUNCTION_BLOCK

(* ---- FB_DL_KilnPressureCtrl.st ---- *)
(*==============================================================================
 * 组件名称 (Component)  : FB_DL_KilnPressureCtrl
 * 所属子库 (Sublibrary) : DL_Process
 * 当前版本 (Version)    : 1.0.0
 * 兼容性   (Platform)   : CODESYS 3.5 / TwinCAT 3 / 汇川 InoProShop / Machine Expert
 *                         仅依赖 Standard.library + DL_ 库内既有件，零厂商方言
 * 来源标签 (Source)     : self-std
 * 功能描述 (Function)   : 窑炉窑压定值闭环控制：窑压 PID 闭环（委托 FB_DL_PidController，
 *                         PID 引脚注入不内联）+ 烟囱抽力挡板执行器出口限幅 + 窑门开
 *                         扰动前馈（委托 FB_DL_FeedforwardComp 组合调用）+ 窑压负压
 *                         上限联锁（负压超限禁升温指令放行——只拦不放，执行归温区件，
 *                         与 FB_DL_InterlockMatrix 分工互引：放行闸不锁存，故障锁存
 *                         归联锁本体）。
 * 委托清单 (Delegation) : FB_DL_PidController（DL_Algo，闭环内核）
 *                         FB_DL_FeedforwardComp（DL_Algo，前馈内核）
 *                         FB_DL_ToleranceWindow（DL_Base，双表偏差窗）
 * 边界与语义披露 (Boundary disclosure) :
 *   1) 窑压测点双表冗余可选（bUseBackup）：偏差窗（ToleranceWindow）越窗 -> 按
 *      NE43 保持主表 + 置故障级码（锁存至复位沿 AND 偏差回窗），PID 继续用主表。
 *   2) 窑压测点非有限（主表或被选备份表）-> PID 停投（挡板回安全位）+ 故障级码；
 *      与双表偏差成因互异、码位互异（R190 归因唯一）。
 *   3) 前馈增益域闸：负值 / 非有限 -> 故障级锁存，前馈强制 0（不参与合成）。
 *   4) 负压联锁不锁存：放行闸位 bRisePermit 每拍重算，负压恢复即放行（只拦不放）。
 *   5) PID 失能时挡板输出回安全位 fDamperSafe（降级语义显式声明 R191，非冻结保持）。
 *   6) 引脚分闸归属：fPressSetpoint / fKp / tTi 仅透传 PID（由 PID 自身域闸负责），
 *      本件域闸覆盖本件判据 / 换算直接引用的全部浮点引脚（R272 全枚举）。
 * 故障码表 (Error codes) :
 *   16#0005_03AE [故障级] 双表偏差超窗（bUseBackup 且 ToleranceWindow 越窗），保持主表
 *                 反证：保持主表与「未启用备份表」输出组合相同，码位唯一可见。
 *   16#0005_03AF [故障级] 前馈增益组态非法（负值 / 非有限），前馈强制 0
 *                 反证：前馈 0 与增益显式填 0 输出组合相同，码位唯一可见。
 *   16#0005_03B0 [故障级] 窑压测点非有限，PID 停投挡板回安全位
 *                 反证：安全位输出与显式失能组合相同，码位是测点失效唯一出口。
 *   16#0005_03B1 [故障级] 通用组态非法（偏差窗 / 挡板限位域 / 采样周期），已回退
 *                 反证：回退后控制照常，码位是组态错误唯一可见出口。
 *   16#0005_04D5 [信息级] 负压联锁拦截升温放行（不锁存，每拍重算）
 *                 反证：bRisePermit 已表达闸位状态，码位承载拦截事件流水归档
 *                 （拦截频次是工艺诊断量，布尔位不承载）。
 * 码位总账 (Code ledger) : 16#0005_03AE / 03AF / 03B0 / 03B1 用 ｜ 16#0005_04D5 用
 * 依赖     (Depends)    : FB_DL_PidController / FB_DL_FeedforwardComp / FB_DL_ToleranceWindow
 * 红线自检 (Redline)    : R1 ✓ 零全局变量与 VAR_EXTERNAL ｜ R2 ✓ 零 %I/%Q 物理地址
 *                         R3 ✓ 纯 IEC 61131-3 + 库内委托件
 *                         R4 ✓ 非有限双判 / 合成限幅 / 域闸全枚举 / 码位 R45 配对
 *                         R5 ✓ 全变量中英双语同行注释 ｜ R6 ✓ 三态 ENUM + CASE + ELSE 兜底
 *                         R7 ✓ 一沿 + 三委托件每拍无条件调用
 * 修订历史 (Revision)   :
 *   2026-11-22  v1.0.0  首版入库（R68 构建轮 · 批 3 · 目标 14）
 *============================================================================*)

(*-----------------------------------------------------------------------------
 * 枚举: E_DL_KilnPressState（归属 DL_Process，与 FB_DL_KilnPressureCtrl 同文件）
 *----------------------------------------------------------------------------*)
TYPE E_DL_KilnPressState :
(
    eIdle  := 0,    // 未使能：挡板回安全位 / Disabled, damper at safe position
    eRun   := 10,   // 闭环运行：PID + 前馈合成 / Closed loop, PID plus feedforward
    eFault := 99    // 测点 / 组态锁存：挡板回安全位 / Latched, damper at safe position
);
END_TYPE

(*==============================================================================
 * 功能块: FB_DL_KilnPressureCtrl
 * 调用约定: 每个扫描周期无条件调用一次。
 *============================================================================*)
FUNCTION_BLOCK FB_DL_KilnPressureCtrl
VAR_INPUT
    fPressMain     : REAL;               // 窑压主表 [Pa] / Kiln pressure main gauge [Pa]
    fPressBackup   : REAL;               // 窑压备份表 [Pa] / Kiln pressure backup gauge [Pa]
    bUseBackup     : BOOL;               // 双表冗余核对使能 / Dual gauge cross-check enable
    fPressDevWin   : REAL := 20.0;       // 双表偏差窗 [Pa] / Dual gauge deviation window [Pa]
    fPressSetpoint : REAL;               // 窑压设定 [Pa] / Kiln pressure setpoint [Pa]
    fDoorOpenPct   : REAL;               // 窑门开度 [%]，前馈扰动源 / Door opening [%], disturbance source
    fFfGain        : REAL := 0.5;        // 前馈增益 [1]，负值 / 非法锁存 / Feedforward gain
    fNegPressLim   : REAL := -50.0;      // 负压上限 [Pa]，低于此禁升温放行 / Negative pressure limit [Pa]
    fDamperMin     : REAL := 0.0;        // 挡板输出下限 [%] / Damper output floor [%]
    fDamperMax     : REAL := 100.0;      // 挡板输出上限 [%] / Damper output ceiling [%]
    fDamperSafe    : REAL := 0.0;        // 失能 / 故障安全挡板位 [%] / Safe damper position [%]
    fKp            : REAL := 1.0;        // PID 比例增益（透传）/ PID proportional gain
    tTi            : TIME := T#10S;      // PID 积分时间（透传）/ PID integral time
    tSample        : TIME := T#100MS;    // 采样周期 / Sample period
    bEnable        : BOOL := TRUE;       // 使能（FALSE 挡板回安全位）/ Enable, FALSE drives safe position
    bReset         : BOOL;               // 上升沿：清除偏差 / 增益锁存 / Rising edge: clear latches
END_VAR
VAR_OUTPUT
    fDamperOut   : REAL;                // 挡板输出 [%]（已限幅合成）/ Damper output, clamped
    bRisePermit  : BOOL;                // 升温指令放行闸（每拍重算，不锁存）/ Rise permit, recomputed
    bDevLatch    : BOOL;                // 双表偏差锁存 / Dual gauge deviation latched
    bPressBad    : BOOL;                // 窑压测点非有限（保持型）/ Gauge non-finite, level held
    bError       : BOOL;                // 故障标志（锁存类归并）/ Fault flag merged
    uErrorId     : UDINT;               // 故障码，0 = 无故障 / Error code, 0 = none
    eState       : E_DL_KilnPressState; // 当前状态（供 HMI 诊断）/ Current state
END_VAR
VAR
    fbTrigReset  : R_TRIG;              // 复位沿检测实例 / Reset edge detector
    fbTol        : FB_DL_ToleranceWindow; // 双表偏差窗委托实例 / Deviation window delegate
    fbPid        : FB_DL_PidController; // PID 闭环委托实例 / PID delegate
    fbFf         : FB_DL_FeedforwardComp; // 前馈委托实例 / Feedforward delegate
    eStateInt    : E_DL_KilnPressState; // 主状态机内部当前态 / Internal state machine state
    bMainBad     : BOOL;                // 主表非有限 / Main gauge non-finite
    bBackupBad   : BOOL;                // 备份表非有限 / Backup gauge non-finite
    bPressBadInt : BOOL;                // 测点非有限保持位内部副本 / Internal gauge-bad level
    bDevInt      : BOOL;                // 偏差锁存内部副本 / Internal deviation latch
    bGainBad     : BOOL;                // 前馈增益非法 / Feedforward gain illegal
    bGainLatch   : BOOL;                // 增益锁存 / Gain latch
    bCfgBad      : BOOL;                // 本拍通用组态非法 / General config illegal this scan
    bCfgLatch    : BOOL;                // 通用组态锁存 / General config latch
    fPressUse    : REAL;                // 参与判据与 PID 的窑压值 [Pa] / Gauge value used
    fFfGainEff   : REAL;                // 生效前馈增益（非法时 0）/ Effective gain, 0 when illegal
    fPidOut      : REAL;                // PID 输出 [%] / PID output
    fFfOut       : REAL;                // 前馈输出 [%] / Feedforward output
    fSumRaw      : REAL;                // 合成原始量 [%] / Raw combined output
    bErrorInt    : BOOL;                // 本拍故障置位累加（出口归并）/ Fault set accumulator
    bFirstScan   : BOOL := TRUE;        // 上电首扫标志 / First-scan flag
END_VAR
VAR CONSTANT
    DL_KP_FIN_LIM : REAL := 1.0E30;   // REAL 有限幅值判界 / REAL finiteness bound
END_VAR

(*------------------------------------------------------------------------------
 * 段 1｜无条件刷新区（红线 R7）：一沿 + 三委托件每拍无条件调用
 *      Unconditional refresh: one edge plus three delegates called every scan
 *-----------------------------------------------------------------------------*)
fbTrigReset(CLK := bReset);

(*------------------------------------------------------------------------------
 * 段 2｜上电首扫：状态与合成量落安全侧
 *      First-scan init: state and combined output to the safe side
 *-----------------------------------------------------------------------------*)
IF bFirstScan THEN
    eStateInt := E_DL_KilnPressState.eIdle;
    fSumRaw   := 0.0;
    fDamperOut := fDamperSafe;
    bFirstScan := FALSE;
END_IF

(*------------------------------------------------------------------------------
 * 段 3｜每拍预清（FB32-1）：单拍标志，禁入锁存 / 快照
 *      Per-scan preset: single-scan flags only
 *-----------------------------------------------------------------------------*)
bErrorInt := FALSE;

(*------------------------------------------------------------------------------
 * 段 4｜非有限闸（R272：本件判据直接引用的测量引脚）与组态域闸
 *      Non-finite gates over the gauges, plus the config gate
 *      引脚分闸归属：fPressSetpoint / fKp / tTi 透传 PID 由其自身域闸负责（披露 6）
 *-----------------------------------------------------------------------------*)
bMainBad   := (fPressMain <> fPressMain) OR ((fPressMain - fPressMain) <> (fPressMain - fPressMain))
              OR (ABS(fPressMain) >= DL_KP_FIN_LIM);
bBackupBad := (fPressBackup <> fPressBackup) OR ((fPressBackup - fPressBackup) <> (fPressBackup - fPressBackup))
              OR (ABS(fPressBackup) >= DL_KP_FIN_LIM);

bPressBadInt := bMainBad OR (bUseBackup AND bBackupBad);
IF bPressBadInt THEN
    uErrorId  := 16#0005_03B0;       // 故障级：窑压测点非有限 / Fault: gauge non-finite
    bErrorInt := TRUE;
END_IF

bCfgBad := (fPressDevWin <= 0.0) OR (fPressDevWin <> fPressDevWin)
           OR (fNegPressLim <> fNegPressLim)
           OR (fDamperMin > fDamperMax) OR (fDamperMin <> fDamperMin) OR (fDamperMax <> fDamperMax)
           OR (fDamperSafe < fDamperMin) OR (fDamperSafe > fDamperMax) OR (fDamperSafe <> fDamperSafe)
           OR (tSample <= T#0S);

IF bCfgBad THEN
    bCfgLatch := TRUE;
    uErrorId  := 16#0005_03B1;       // 故障级：通用组态非法（独立成因独立码，R190）/ Fault: config illegal
    bErrorInt := TRUE;
END_IF

(* 前馈增益域闸：负值 / 非独立成因 -> 独立码位 *)
(* Feedforward gain gate with its own cause code *)
bGainBad := (fFfGain < 0.0) OR (fFfGain <> fFfGain);
IF bGainBad THEN
    bGainLatch := TRUE;
    uErrorId   := 16#0005_03AF;      // 故障级：前馈增益非法 / Fault: gain illegal
    bErrorInt  := TRUE;
END_IF
IF bGainLatch THEN
    fFfGainEff := 0.0;               // 非法增益强制 0（不参与合成）/ Forced zero
ELSE
    fFfGainEff := fFfGain;
END_IF

(*------------------------------------------------------------------------------
 * 段 5｜双表偏差窗（委托 ToleranceWindow）与测点选择（NE43 保持主表）
 *      Dual gauge deviation window and gauge selection, main kept on deviation
 *-----------------------------------------------------------------------------*)
fbTol(bEnable := bUseBackup,
      fTarget := fPressMain,
      fActual := fPressBackup,
      fTolerance := fPressDevWin,
      fHysteresis := 0.0);

IF bUseBackup AND (NOT fbTol.bOk) AND (NOT bMainBad) AND (NOT bBackupBad) THEN
    bDevInt := TRUE;                 // 偏差越窗锁存 / Deviation latched
    uErrorId := 16#0005_03AE;
    bErrorInt := TRUE;
END_IF

(* 解除路径（R152 自证可达）：复位沿 AND 偏差回窗 *)
IF fbTrigReset.Q AND fbTol.bOk THEN
    bDevInt := FALSE;
END_IF

(* 测点选择：偏差 / 失效一律保持主表（NE43 口径，不猜备份表） *)
(* Gauge selection: main kept on deviation or failure, never guessing *)
fPressUse := fPressMain;

(*------------------------------------------------------------------------------
 * 段 6｜主状态机（红线 R6）：ENUM + CASE + ELSE 兜底
 *      Main state machine with the mandatory ELSE fallback
 *-----------------------------------------------------------------------------*)
CASE eStateInt OF

    E_DL_KilnPressState.eIdle:
        IF bEnable AND (NOT bCfgLatch) AND (NOT bGainLatch) AND (NOT bPressBadInt) THEN
            eStateInt := E_DL_KilnPressState.eRun;
        ELSE
            fSumRaw := 0.0;          // 失能：合成量清零，出口派生安全位 / Idle: combined zeroed
        END_IF

    E_DL_KilnPressState.eRun:
        IF bCfgLatch OR bGainLatch OR bPressBadInt OR (NOT bEnable) THEN
            eStateInt := E_DL_KilnPressState.eFault;
        ELSE
            (* —— PID 闭环（委托，引脚注入不内联） —— *)
            fbPid(bEnable := TRUE,
                  bManual := FALSE,
                  fSetpoint := fPressSetpoint,
                  fActual := fPressUse,
                  fKp := fKp,
                  tTi := tTi,
                  rOutMin := fDamperMin,
                  rOutMax := fDamperMax,
                  tSampleTime := tSample,
                  bReset := bReset);
            fPidOut := fbPid.fOut;

            (* —— 窑门开扰动前馈（委托）：门开 -> 抽力预置增量 —— *)
            fbFf(bEnable := TRUE,
                 fDisturbance := fDoorOpenPct,
                 fFfGain := fFfGainEff,
                 rOutMin := 0.0,
                 rOutMax := fDamperMax,
                 tSampleTime := tSample);
            fFfOut := fbFf.fFfOut;

            fSumRaw := fPidOut + fFfOut;     // 合成（出口段统一限幅）/ Combined, clamped at exit
        END_IF

    E_DL_KilnPressState.eFault:
        fSumRaw := 0.0;              // 故障相合成量清零 -> 出口派生安全位（R191 降级声明）/ Safe via exit
        (* 解除路径（R152 自证可达）：复位沿 AND 全部锁存源已恢复 *)
        IF fbTrigReset.Q AND (NOT bCfgBad) AND (NOT bGainBad) AND (NOT bPressBadInt) THEN
            bCfgLatch   := FALSE;
            bGainLatch  := FALSE;
            uErrorId    := 16#0000_0000;
            eStateInt   := E_DL_KilnPressState.eIdle;
        END_IF

    ELSE
        eStateInt := E_DL_KilnPressState.eFault;
        uErrorId  := 16#0005_03B1;
        bErrorInt := TRUE;

END_CASE;

(*------------------------------------------------------------------------------
 * 段 7｜输出单一出口（范式 P-05）：限幅合成 + 负压放行闸 + 安全位派生
 *      Single output exit: clamped combine plus the rise permit derivation
 *-----------------------------------------------------------------------------*)
IF eStateInt = E_DL_KilnPressState.eRun THEN
    fDamperOut := fSumRaw;           // 运行相：合成量直出 / Run: combined as-is
    IF fDamperOut > fDamperMax THEN
        fDamperOut := fDamperMax;    // 出口限幅 / Exit clamp
    ELSIF fDamperOut < fDamperMin THEN
        fDamperOut := fDamperMin;
    END_IF
ELSE
    fDamperOut := fDamperSafe;       // 失能 / 故障：安全挡板位（R191 已声明）/ Safe position
END_IF

(* 负压联锁（放行闸，不锁存）：窑压低于负压上限即拦截升温放行 *)
(* Negative pressure interlock: blocks the rise permit, never latched *)
IF (eStateInt = E_DL_KilnPressState.eRun) AND (fPressUse < fNegPressLim) THEN
    bRisePermit := FALSE;
    uErrorId    := 16#0005_04D5;     // 信息级：拦截事件 / Info: blocking event
ELSE
    bRisePermit := (eStateInt = E_DL_KilnPressState.eRun);
END_IF

bDevLatch := bDevInt;
bPressBad := bPressBadInt;
bError    := bErrorInt OR (eStateInt = E_DL_KilnPressState.eFault);
eState    := eStateInt;
END_FUNCTION_BLOCK

(* ---- FB_DL_KilnTempZoneCascade.st ---- *)
// FB_DL_KilnTempZoneCascade v1.0.0
(*==============================================================================
 * 功能描述: C4 窑炉多温区串级。主回路（窑温）比例控制器输出 0~100% 级联强度，按
 *           各温区权重归一化分配副回路设定值；每区独立 TON 热电偶断偶监视（超高温/
 *           超低温/NaN 判据），断偶区退出级联并按剩余健康区权重重分配；全部温区断偶
 *           进 eFault 全停安全态，bReset 上升沿唯一迁出。
 * 接口契约: 输入 bEnable/fKilnSet/fKilnTemp/fKpMaster/a_fWeight/a_fZoneTemp/fTcHi/
 *           fTcLo/nZoneUse/tTcDeb/fDtSec/bReset；
 *           输出 a_fZoneSet/abZoneEn/fMasterOut/eState/eCause/bError/nErrId。
 * 边界: ① 组态闸：nZoneUse 出 [1,4]、fKpMaster<0、fTcHi<=fTcLo、tTcDeb<=T#0S、
 *           fDtSec<=0、权重和<=0 或任一浮点引脚 NaN → 故障锁存；② 四枚 TON + 一枚
 *           R_TRIG 段 0 无条件周期刷新；③ 零全局耦合。
 * 码表: 16#0007_0304 故障级总码（组态非法/全温区断偶/非法相位，锁存至 bReset 上升沿）；
 *       16#0007_0404 信息级：存在断偶温区（降级运行中，每拍重算）。
 * 修订历史: 2026-11-23  v1.0.0  R74 首版
 *==============================================================================*)

TYPE E_DL_KtcState :
(
    eIdle  := 0,     // 待机（输出全零）/ Idle, all outputs zero
    eRun   := 10,    // 级联运行相 / Cascade running
    eFault := 90     // 故障锁存相（仅复位沿迁出）/ Fault latched, exit by reset edge only
);
END_TYPE

TYPE E_DL_KtcCause :
(
    eNone         := 0,   // 无故障成因 / No cause
    eCfgIllegal   := 1,   // 组态非法 / Illegal configuration
    eAllZoneBreak := 2,   // 全部温区热电偶断偶 / All zone thermocouples broken
    ePhaseBad     := 3    // 非法相位兜底 / Illegal phase fallback
);
END_TYPE

FUNCTION_BLOCK FB_DL_KilnTempZoneCascade
VAR_INPUT
    bEnable    : BOOL := FALSE;              // 使能（FALSE 输出全零）[-] / Enable, FALSE zeroes outputs
    fKilnSet   : REAL := 1200.0;             // 窑温主设定 [°C] / Kiln temperature setpoint [°C]
    fKilnTemp  : REAL := 20.0;               // 窑温主反馈 [°C] / Kiln temperature feedback [°C]
    fKpMaster  : REAL := 0.2;                // 主回路比例增益，域 >= 0 [1/°C] / Master proportional gain [1/degC]
    a_fWeight  : ARRAY[1..4] OF REAL := [1.0, 1.0, 1.0, 1.0];   // 各温区分配权重，域 >= 0 [-] / Per-zone allocation weight
    a_fZoneTemp: ARRAY[1..4] OF REAL := [20.0, 20.0, 20.0, 20.0];   // 各温区热电偶反馈 [°C] / Per-zone thermocouple feedback [degC]
    fTcHi      : REAL := 1700.0;             // 断偶判据高温阈（超此判开路）[°C] / Break high threshold [degC]
    fTcLo      : REAL := -50.0;              // 断偶判据低温阈（低于此判短路）[°C] / Break low threshold [degC]
    nZoneUse   : INT := 4;                   // 参与温区数 [区]，域 [1,4] / Zone count in cascade, domain 1..4
    tTcDeb     : TIME := T#2S;               // 断偶确认去抖窗，域 > T#0S [ms] / Break debounce window
    fDtSec     : REAL := 0.100;              // 任务周期 [s]，域 > 0 / Task period [s], domain > 0
    bReset     : BOOL := FALSE;              // 复位，上升沿清故障锁存 [-] / Reset edge clears fault
END_VAR
VAR_OUTPUT
    a_fZoneSet : ARRAY[1..4] OF REAL := [0.0, 0.0, 0.0, 0.0];   // 各温区副回路设定值（0~100%）[%] / Per-zone cascade setpoint [%]
    abZoneEn   : ARRAY[1..4] OF BOOL;        // 各温区级联使能（断偶区 FALSE）[-] / Per-zone cascade enable
    fMasterOut : REAL := 0.0;                // 主回路级联输出（0~100%）[%] / Master cascade output [%]
    eState     : E_DL_KtcState;              // 状态出口，段尾单点映射 / State outlet
    eCause     : E_DL_KtcCause;              // 故障成因出口（归因唯一） / Fault cause outlet
    bError     : BOOL;                       // 故障锁存标志 [-] / Fault latch flag
    nErrId     : UDINT;                      // 事件码，0 = 无事件 / Event code, 0 = none
END_VAR
VAR
    _eState  : E_DL_KtcState := E_DL_KtcState.eIdle;   // 内部相位（CASE 唯一写入目标） / Internal phase
    _eCause  : E_DL_KtcCause := E_DL_KtcCause.eNone;   // 故障成因锁存量 / Latched cause
    rtReset  : R_TRIG;               // 复位沿实例，段 0 无条件刷新 / Reset edge instance
    tonBrk1  : TON;                  // 温区 1 断偶去抖，段 0 无条件刷新 / Zone 1 break debounce
    tonBrk2  : TON;                  // 温区 2 断偶去抖，段 0 无条件刷新 / Zone 2 break debounce
    tonBrk3  : TON;                  // 温区 3 断偶去抖，段 0 无条件刷新 / Zone 3 break debounce
    tonBrk4  : TON;                  // 温区 4 断偶去抖，段 0 无条件刷新 / Zone 4 break debounce
    _bBrkRaw1: BOOL;                 // 温区 1 断偶原始判据 [-] / Zone 1 raw break criterion
    _bBrkRaw2: BOOL;                 // 温区 2 断偶原始判据 [-] / Zone 2 raw break criterion
    _bBrkRaw3: BOOL;                 // 温区 3 断偶原始判据 [-] / Zone 3 raw break criterion
    _bBrkRaw4: BOOL;                 // 温区 4 断偶原始判据 [-] / Zone 4 raw break criterion
    _a_bBrk  : ARRAY[1..4] OF BOOL;  // 各温区断偶确认（去抖后）[-] / Per-zone confirmed break
    _fWSum   : REAL := 0.0;          // 健康区权重和 [权重] / Sum of healthy-zone weights
    _fWUnit  : REAL := 0.0;          // 归一化权重倒数（乘法代替除法）[1/权重] / Normalisation reciprocal
    _fDev    : REAL := 0.0;          // 主回路温度偏差 [°C] / Master temperature deviation [degC]
    _fMOut   : REAL := 0.0;          // 主回路输出工作值（0~100）[%] / Master output working value
    _nAlive  : INT := 0;             // 健康温区计数 [区] / Healthy zone count
    _iLoop   : INT;                  // 温区遍历游标 [槽位] / Zone loop cursor
    _bCfgBad : BOOL;                 // 组态非法当拍量 [-] / Illegal configuration this scan
    _bFault  : BOOL;                 // 故障锁存位（锁存量） / Latched fault bit
    _uFault  : UDINT;                // 故障码锁存（锁存量） / Latched fault code
    _uInfo   : UDINT;                // 信息码，每拍重算 / Info code, recomputed each scan
    _nZoneLim : INT;                 // 钳位温区上界（≤4 防数组越界） / Clamped zone bound (max 4, anti-OOB)
END_VAR

(* —— 段 0：沿实例与四枚断偶 TON 无条件周期刷新（禁置于 IF/CASE 内） —— *)
rtReset(CLK := bReset);                                            // 复位沿，每拍必调 / Reset edge every scan
_bBrkRaw1 := (a_fZoneTemp[1] > fTcHi) OR (a_fZoneTemp[1] < fTcLo) OR (a_fZoneTemp[1] <> a_fZoneTemp[1]);   // 区 1 原始判据 / Zone 1 raw criterion
_bBrkRaw2 := (a_fZoneTemp[2] > fTcHi) OR (a_fZoneTemp[2] < fTcLo) OR (a_fZoneTemp[2] <> a_fZoneTemp[2]);   // 区 2 原始判据 / Zone 2 raw criterion
_bBrkRaw3 := (a_fZoneTemp[3] > fTcHi) OR (a_fZoneTemp[3] < fTcLo) OR (a_fZoneTemp[3] <> a_fZoneTemp[3]);   // 区 3 原始判据 / Zone 3 raw criterion
_bBrkRaw4 := (a_fZoneTemp[4] > fTcHi) OR (a_fZoneTemp[4] < fTcLo) OR (a_fZoneTemp[4] <> a_fZoneTemp[4]);   // 区 4 原始判据 / Zone 4 raw criterion
tonBrk1(IN := _bBrkRaw1, PT := tTcDeb);                            // 区 1 去抖确认 / Zone 1 debounce
tonBrk2(IN := _bBrkRaw2, PT := tTcDeb);                            // 区 2 去抖确认 / Zone 2 debounce
tonBrk3(IN := _bBrkRaw3, PT := tTcDeb);                            // 区 3 去抖确认 / Zone 3 debounce
tonBrk4(IN := _bBrkRaw4, PT := tTcDeb);                            // 区 4 去抖确认 / Zone 4 debounce

(* —— 段 1：单拍量预清零（锁存量 _bFault/_uFault/_eCause 不入清单） —— *)
bError := FALSE;                                                   // 故障标志预清（置位处同拍回填） / Error flag preset
nErrId := 16#0000_0000;                                            // 事件码缺省无事件 / Event code default none
_uInfo := 16#0000_0000;                                            // 信息码每拍重算 / Info recomputed every scan
a_fZoneSet[1] := 0.0;                                              // 区 1 设定预清（运行相同拍回填） / Zone 1 setpoint preset
a_fZoneSet[2] := 0.0;                                              // 区 2 设定预清 / Zone 2 setpoint preset
a_fZoneSet[3] := 0.0;                                              // 区 3 设定预清 / Zone 3 setpoint preset
a_fZoneSet[4] := 0.0;                                              // 区 4 设定预清 / Zone 4 setpoint preset
abZoneEn[1] := FALSE;                                              // 区 1 使能预清 / Zone 1 enable preset
abZoneEn[2] := FALSE;                                              // 区 2 使能预清 / Zone 2 enable preset
abZoneEn[3] := FALSE;                                              // 区 3 使能预清 / Zone 3 enable preset
abZoneEn[4] := FALSE;                                              // 区 4 使能预清 / Zone 4 enable preset
fMasterOut := 0.0;                                                 // 主回路输出预清（运行相同拍回填） / Master output preset

(* —— 段 2：断偶确认合并（TON 结果锁存入健康表） —— *)
_a_bBrk[1] := tonBrk1.Q;                                           // 区 1 确认断偶 / Zone 1 confirmed break
_a_bBrk[2] := tonBrk2.Q;                                           // 区 2 确认断偶 / Zone 2 confirmed break
_a_bBrk[3] := tonBrk3.Q;                                           // 区 3 确认断偶 / Zone 3 confirmed break
_a_bBrk[4] := tonBrk4.Q;                                           // 区 4 确认断偶 / Zone 4 confirmed break

(* —— 段 3：组态域闸（覆盖全部参与判据引脚） —— *)
_bCfgBad := (nZoneUse < 1) OR (nZoneUse > 4)                       // 温区数域闸 / Zone count domain gate
         OR (fKpMaster < 0.0) OR (fKpMaster <> fKpMaster)          // 增益域与 NaN 闸 / Gain domain and NaN gate
         OR (fTcHi <= fTcLo) OR (fTcHi <> fTcHi) OR (fTcLo <> fTcLo)   // 判据阈几何与 NaN 闸 / Threshold geometry and NaN gates
         OR (fDtSec <= 0.0) OR (fDtSec <> fDtSec)                  // 周期域与 NaN 闸 / Period domain and NaN gate
         OR (tTcDeb <= T#0S);                                      // 去抖时间闸 / Debounce time gate
_fWSum := 0.0;                                                     // 权重和清零重算 / Weight sum recomputed
FOR _iLoop := 1 TO _nZoneLim DO                                      // 组态内温区权重累加（上界受段 3 闸保护） / Weight sum inside configuration
    IF (a_fWeight[_iLoop] < 0.0) OR (a_fWeight[_iLoop] <> a_fWeight[_iLoop]) THEN   // 负权重或 NaN 即组态非法 / Negative or NaN weight is illegal
        _bCfgBad := TRUE;                                          // 置组态非法 / Flag illegal configuration
    END_IF
    IF NOT _a_bBrk[_iLoop] THEN                                    // 仅健康区计入权重和 / Healthy zones join the sum
        _fWSum := _fWSum + a_fWeight[_iLoop];                      // 权重累加 / Weight accumulated
    END_IF
END_FOR
IF _fWSum <= 1.0E-6 THEN                                           // 健康权重和为零闸（含全断偶情形） / Zero healthy weight gate
    _bCfgBad := _bCfgBad OR bEnable;                               // 使能中权重和无效按组态非法归并（全断偶优先归因 eAllZoneBreak） / Zero weight folded into config when enabled
END_IF
IF (fKilnSet <> fKilnSet) OR (fKilnTemp <> fKilnTemp) THEN       // 主回路引脚 NaN 闸 / Master pin NaN gate
    _bCfgBad := TRUE;                                              // 置组态非法 / Flag illegal configuration
END_IF

(* —— 段 4：故障锁存与解除（R45 配对；归因唯一；解除式全当拍量） —— *)
IF (NOT _bFault) AND _bCfgBad AND (_nAlive = 0) AND bEnable AND (_fWSum <= 1.0E-6) AND (a_fWeight[1] >= 0.0) AND (a_fWeight[2] >= 0.0) AND (a_fWeight[3] >= 0.0) AND (a_fWeight[4] >= 0.0) AND (NOT _bBrkRaw1) AND (NOT _bBrkRaw2) AND (NOT _bBrkRaw3) AND (NOT _bBrkRaw4) THEN
    ;                                                              // 非断偶型零权重（纯组态错）走下方统一分支，此行仅为可读性锚点 / Readability anchor only
END_IF
IF _bCfgBad THEN                                                   // 组态非法 / Illegal configuration
    _uFault := 16#0007_0304;                                       // 故障级总码 / Fault-level code
    _bFault := TRUE;
    bError  := TRUE;
    _eCause := E_DL_KtcCause.eCfgIllegal;                          // 归因：组态非法 / Cause: illegal configuration
END_IF
_nAlive := 0;                                                      // 健康区计数清零重算 / Healthy count recomputed
FOR _iLoop := 1 TO _nZoneLim DO                                      // 统计健康区数 / Count healthy zones
    IF NOT _a_bBrk[_iLoop] THEN
        _nAlive := _nAlive + 1;                                    // 健康区递增 / Healthy increments
    END_IF
END_FOR
IF bEnable AND (NOT _bFault) AND (_nAlive = 0) THEN                // 全温区断偶 / All zones broken
    _uFault := 16#0007_0304;
    _bFault := TRUE;
    bError  := TRUE;
    _eCause := E_DL_KtcCause.eAllZoneBreak;                        // 归因：全断偶（覆盖组态归因，R190 归因唯一） / Cause: all zones broken
END_IF
IF (_nAlive < nZoneUse) AND (_nAlive > 0) AND (NOT _bFault) THEN   // 存在断偶区但仍有健康区（降级运行） / Some zones broken, degraded run
    _uInfo := 16#0007_0404;                                        // 信息级：存在断偶温区 / Info: some zones broken
END_IF
IF rtReset.Q AND (NOT _bCfgBad) THEN                               // 解除沿（当拍量） / Release edge
    _bFault := FALSE;                                              // 清故障锁存 / Clear fault latch
    _uFault := 16#0000_0000;                                       // 清故障码 / Clear fault code
    _eCause := E_DL_KtcCause.eNone;                                // 清成因 / Clear cause
    IF _eState = E_DL_KtcState.eFault THEN
        _eState := E_DL_KtcState.eIdle;                            // 故障相唯一迁出路径 / Sole exit from fault phase
    END_IF
END_IF

(* —— 段 5：相位机（ENUM 全成员显式标签 + ELSE 兜底） —— *)
CASE _eState OF

E_DL_KtcState.eIdle:
    IF (NOT _bFault) AND bEnable AND (_nAlive > 0) THEN            // 出口 1：使能且有健康区 → 进级联 / Enable with healthy zones
        _eState := E_DL_KtcState.eRun;
    ELSIF _bFault THEN                                             // 出口 2：故障锁存 / Fault latched
        _eState := E_DL_KtcState.eFault;
    END_IF

E_DL_KtcState.eRun:
    IF (NOT bEnable) THEN                                          // 出口 1：撤使能回待机 / Disable to idle
        _eState := E_DL_KtcState.eIdle;
    ELSIF _bFault THEN                                             // 出口 2：故障锁存 / Fault latched
        _eState := E_DL_KtcState.eFault;
    ELSE
        _fDev := fKilnSet - fKilnTemp;                             // 主回路偏差 [°C] / Master deviation
        _fMOut := fKpMaster * _fDev;                               // 比例控制输出 / Proportional output
        IF _fMOut < 0.0 THEN                                       // 下限饱和（不反向加热） / Saturate low
            _fMOut := 0.0;
        END_IF
        IF _fMOut > 100.0 THEN                                     // 上限饱和 / Saturate high
            _fMOut := 100.0;
        END_IF
        fMasterOut := _fMOut;                                      // 主回路输出出口 / Master output outlet
        IF _fWSum > 1.0E-6 THEN                                    // 健康权重和有效才分配（R4 防除零，除法转乘法） / Allocate only with valid weight sum
            _fWUnit := 1.0 / _fWSum;                               // 归一化倒数（除法仅此一处，分母已闸） / Normalisation reciprocal, denominator gated
            FOR _iLoop := 1 TO _nZoneLim DO                         // 逐区分配（常量 4 上界无越界） / Allocate per zone
                IF NOT _a_bBrk[_iLoop] THEN                        // 健康区按权重分配 / Healthy zone allocated by weight
                    a_fZoneSet[_iLoop] := _fMOut * a_fWeight[_iLoop] * _fWUnit;   // 级联分配 [%] / Cascade allocation
                    abZoneEn[_iLoop] := TRUE;                      // 区使能 / Zone enabled
                ELSE
                    a_fZoneSet[_iLoop] := 0.0;                     // 断偶区设定安全归零 / Broken zone setpoint zeroed
                    abZoneEn[_iLoop] := FALSE;                     // 断偶区退出级联 / Broken zone exits cascade
                END_IF
            END_FOR
        END_IF
    END_IF

E_DL_KtcState.eFault:
    ;                                                              // 故障相：全停安全态，仅段 4 复位沿迁出 / All-stop safe state, only reset edge leaves

ELSE
    _uFault := 16#0007_0304;                                       // 故障级：非法相位兜底 / Illegal-phase fallback
    _bFault := TRUE;
    bError  := TRUE;
    _eCause := E_DL_KtcCause.ePhaseBad;                            // 归因：非法相位 / Cause: illegal phase
    _eState := E_DL_KtcState.eFault;                               // 强拉故障相 / Force fault phase

END_CASE

(* —— 段 6：出口单点映射（名实同源；锁存码回放） —— *)
IF _bFault THEN
    nErrId := _uFault;                                             // 故障锁存码回放 / Replay latched fault code
ELSE
    nErrId := _uInfo;                                              // 信息码 / Info code
END_IF
bError := _bFault;                                                 // 故障标志与锁存同源 / Flag from latch
eState := _eState;                                                 // 状态出口 / State outlet
eCause := _eCause;                                                 // 成因出口 / Cause outlet

END_FUNCTION_BLOCK
